// Упакованный канал: подготовка payload -> CommandSeq -> Result -> Ack.
udiGeometryRequest := GVL_HMI.udiGeometryCommandSeq;
xGeometryRequestFresh := FALSE;
IF (udiGeometryRequest <> UDINT#0) AND (udiGeometryRequest <> GVL_HMI.udiGeometryAckSeq) THEN
	stGeometryRequest := GVL_HMI.stGeometryRequest;
	GVL_HMI.uiGeometryResult := UINT#2;
	IF NOT IsHmiCommandFresh(udiIssuedAtMs := GVL_HMI.udiGeometryIssuedAtMs) THEN
		GVL_HMI.uiGeometryResult := UINT#4;
	ELSIF xHmiConnectionAlive THEN
		xGeometryRequestFresh := TRUE;
		IF (stGeometryRequest.uiAction = UINT#8) AND (stGeometryRequest.uiMachine >= UINT#1)
		AND (stGeometryRequest.uiMachine <= UINT#3) THEN
			uiGeometryMachine := stGeometryRequest.uiMachine;
			IF GVL_GEOMETRY_CONTROL.axCallAllowed[uiGeometryMachine] THEN
				IF GVL_GEOMETRY_CONTROL.astCalls[uiGeometryMachine].uiState = UINT#1 THEN
					stGeometryCall := GVL_GEOMETRY_CONTROL.astCalls[uiGeometryMachine];
				ELSE
					GVL_GEOMETRY_CONTROL.udiNextCallId := GVL_GEOMETRY_CONTROL.udiNextCallId + UDINT#1;
					IF GVL_GEOMETRY_CONTROL.udiNextCallId = UDINT#0 THEN GVL_GEOMETRY_CONTROL.udiNextCallId := UDINT#1; END_IF;
					stGeometryCall := stGeometryEmptyCall;
					stGeometryCall.udiId := GVL_GEOMETRY_CONTROL.udiNextCallId;
					stGeometryCall.uiMachine := uiGeometryMachine;
					stGeometryCall.uiProductType := GVL_MULTI_TYPE.Config.auiMachineType[uiGeometryMachine];
				END_IF;
				stGeometryCall.xForced := TRUE; stGeometryCall.uiState := UINT#1;
				GVL_GEOMETRY_CONTROL.astCalls[uiGeometryMachine] := stGeometryCall;
				GVL_GEOMETRY_CONTROL.auiActiveCount[uiGeometryMachine] := UINT#0;
				F_GEOMETRY_EVENT(Call := stGeometryCall); GVL_HMI.uiGeometryResult := UINT#1;
			END_IF;
		ELSIF (stGeometryRequest.uiAction = UINT#12) AND (stGeometryRequest.uiMachine >= UINT#1)
		AND (stGeometryRequest.uiMachine <= UINT#3) THEN
			uiGeometryMachine := stGeometryRequest.uiMachine;
			IF GVL_GEOMETRY_CONTROL.axCancelAllowed[uiGeometryMachine] THEN
				GVL_GEOMETRY_CONTROL.astCalls[uiGeometryMachine].uiState := UINT#6;
				F_GEOMETRY_EVENT(Call := GVL_GEOMETRY_CONTROL.astCalls[uiGeometryMachine]); GVL_HMI.uiGeometryResult := UINT#1;
			END_IF;
		ELSIF (stGeometryRequest.uiAction = UINT#9) AND GVL_GEOMETRY_CONTROL.xAutoChangeAllowed
		AND (stGeometryRequest.udiValue <= UDINT#1) THEN
			GVL_GEOMETRY_CONTROL.xAutoEnabled := stGeometryRequest.udiValue = UDINT#1;
			GVL_HMI.uiGeometryResult := UINT#1;
		ELSIF (stGeometryRequest.uiAction = UINT#10) AND GVL_GEOMETRY_CONTROL.xAutoChangeAllowed
		AND (stGeometryRequest.uiMachine <= UINT#3) AND (stGeometryRequest.udiValue >= UDINT#1)
		AND (stGeometryRequest.udiValue <= UDINT#10000) THEN
			FOR uiGeometryMachine := UINT#1 TO UINT#3 DO
				IF (stGeometryRequest.uiMachine = UINT#0) OR (stGeometryRequest.uiMachine = uiGeometryMachine) THEN
					GVL_GEOMETRY_CONTROL.auiPeriod[uiGeometryMachine] := UDINT_TO_UINT(stGeometryRequest.udiValue);
				END_IF;
			END_FOR;
			GVL_HMI.uiGeometryResult := UINT#1;
		ELSIF (stGeometryRequest.uiAction = UINT#16) AND GVL_GEOMETRY_CONTROL.xSettingsAllowed THEN
			CASE stGeometryRequest.uiMachine OF
				UINT#1: IF stGeometryRequest.udiValue <= UDINT#1 THEN GVL_GEOMETRY_CONTROL.xWaitWhenOccupied := stGeometryRequest.udiValue = UDINT#1; GVL_HMI.uiGeometryResult := UINT#1; END_IF;
				UINT#2: IF (stGeometryRequest.udiValue >= UDINT#100) AND (stGeometryRequest.udiValue <= UDINT#600000) THEN GVL_GEOMETRY_CONTROL.tTransportTimeout := UDINT_TO_TIME(stGeometryRequest.udiValue); GVL_HMI.uiGeometryResult := UINT#1; END_IF;
				UINT#3: IF (stGeometryRequest.udiValue >= UDINT#100) AND (stGeometryRequest.udiValue <= UDINT#60000) THEN GVL_GEOMETRY_CONTROL.tDriveFeedbackTimeout := UDINT_TO_TIME(stGeometryRequest.udiValue); GVL_HMI.uiGeometryResult := UINT#1; END_IF;
				UINT#4: IF (stGeometryRequest.udiValue >= UDINT#100) AND (stGeometryRequest.udiValue <= UDINT#10000) THEN GVL_GEOMETRY_CONTROL.tResetPulse := UDINT_TO_TIME(stGeometryRequest.udiValue); GVL_HMI.uiGeometryResult := UINT#1; END_IF;
				UINT#5: IF (stGeometryRequest.udiValue >= UDINT#1000) AND (stGeometryRequest.udiValue <= UDINT#3600000) THEN GVL_GEOMETRY_CONTROL.tWaitWarningTimeout := UDINT_TO_TIME(stGeometryRequest.udiValue); GVL_HMI.uiGeometryResult := UINT#1; END_IF;
			END_CASE;
		ELSIF (stGeometryRequest.uiStation >= UINT#1) AND (stGeometryRequest.uiStation <= UINT#2) THEN
			uiGeometry := stGeometryRequest.uiStation;
			IF (stGeometryRequest.uiAction >= UINT#1) AND (stGeometryRequest.uiAction <= UINT#7) THEN
				GVL_GEOMETRY_CONTROL.auiAction[uiGeometry] := stGeometryRequest.uiAction;
			ELSIF (stGeometryRequest.uiAction = UINT#11) AND GVL_GEOMETRY_CONTROL.xSupported
			AND GVL_POINT_MANAGER.PointManager.Diag.xXLimitValid
			AND GVL_POINT_MANAGER.PointManager.Diag.xYLimitValid
			AND GVL_POINT_MANAGER.PointManager.Diag.xZLimitValid THEN
				stGeometryConfig := stGeometryRequest.Config;
				stGeometryConfig.lrChangeZ := stGeometryConfig.lrSafeZ;
				xGeometryConfigValid := (stGeometryConfig.lrSpeedFactor >= 0.1) AND (stGeometryConfig.lrSpeedFactor <= 1.0)
					AND (stGeometryConfig.lrSafeZ < 0.0) AND (stGeometryConfig.lrSafeZ >= -10000.0)
					AND (stGeometryConfig.lrX >= GVL_POINT_MANAGER.PointManager.Diag.lrX_MinLimit)
					AND (stGeometryConfig.lrX <= GVL_POINT_MANAGER.PointManager.Diag.lrX_MaxLimit)
					AND (stGeometryConfig.lrY >= GVL_POINT_MANAGER.PointManager.Diag.lrY_MinLimit)
					AND (stGeometryConfig.lrY <= GVL_POINT_MANAGER.PointManager.Diag.lrY_MaxLimit)
					AND (stGeometryConfig.lrZ >= GVL_POINT_MANAGER.PointManager.Diag.lrZ_MinLimit)
					AND (stGeometryConfig.lrZ <= GVL_POINT_MANAGER.PointManager.Diag.lrZ_MaxLimit)
					AND ((stGeometryConfig.lrZ + stGeometryConfig.lrSafeZ) >= GVL_POINT_MANAGER.PointManager.Diag.lrZ_MinLimit);
				IF xGeometryConfigValid THEN
					stGeometryConfig.xConfigured := TRUE;
					IF GVL_CELL_SETTINGS.eTestEnvironment = E_CELL_TEST_ENVIRONMENT.NORMAL THEN GVL_GEOMETRY_CONTROL.astConfig[uiGeometry] := stGeometryConfig;
					ELSE GVL_GEOMETRY_CONTROL.astSimulationConfig[uiGeometry] := stGeometryConfig; END_IF;
					GVL_GEOMETRY_CONTROL.astActiveConfig[uiGeometry] := stGeometryConfig; GVL_HMI.uiGeometryResult := UINT#1;
				END_IF;
			ELSIF (stGeometryRequest.uiAction = UINT#13) AND GVL_GEOMETRY_CONTROL.astStatus[uiGeometry].xPointWriteAllowed
			AND GVL_HMI.xPointEditorCaptureAllowed THEN
				GVL_HMI.stGeometryCapture := GVL_GEOMETRY_CONTROL.astActiveConfig[uiGeometry];
				GVL_HMI.stGeometryCapture.lrX := lrRobotActualX; GVL_HMI.stGeometryCapture.lrY := lrRobotActualY;
				GVL_HMI.stGeometryCapture.lrZ := lrRobotActualZ; GVL_HMI.uiGeometryResult := UINT#1;
			ELSIF ((stGeometryRequest.uiAction = UINT#14) OR (stGeometryRequest.uiAction = UINT#15))
			AND GVL_CELL_SETTINGS.xErrorSimulationEnabled
			AND (GVL_CELL_SETTINGS.eTestEnvironment = E_CELL_TEST_ENVIRONMENT.SIMULATION)
			AND GVL_GEOMETRY_CONTROL.xSupported THEN
				GVL_GEOMETRY_CONTROL.axSimulationAlarm[uiGeometry] := stGeometryRequest.uiAction = UINT#14;
				GVL_HMI.uiGeometryResult := UINT#1;
			END_IF;
		END_IF;
	END_IF;
END_IF;

FOR uiGeometry := UINT#1 TO UINT#2 DO
	xGeometryStopAttempt := FALSE;
	IF (GVL_HMI.audiGeometryStopSeq[uiGeometry] <> UDINT#0)
	AND (GVL_HMI.audiGeometryStopSeq[uiGeometry] <> GVL_HMI.audiGeometryStopAck[uiGeometry]) THEN
		GVL_GEOMETRY_CONTROL.auiAction[uiGeometry] := UINT#6;
		xGeometryStopAttempt := TRUE;
		GVL_HMI.audiGeometryStopAck[uiGeometry] := GVL_HMI.audiGeometryStopSeq[uiGeometry];
	END_IF;
	IF GVL_CELL_SETTINGS.eTestEnvironment <> E_CELL_TEST_ENVIRONMENT.NORMAL THEN
		GEOMETRY_SIM[uiGeometry](xInitialize := xGeometryEnvironmentChanged OR xTestInitializePulse,
			xRun := GEOMETRY[uiGeometry].xRunOutput, xReset := GEOMETRY[uiGeometry].xResetOutput,
			xDeposited := GVL_GEOMETRY_CONTROL.astSignals[uiGeometry].xDeposited,
			udiPartId := GVL_GEOMETRY_CONTROL.astSignals[uiGeometry].Call.udiId,
			xRemove := GEOMETRY[uiGeometry].xSimulationEmptyConfirmed,
			xAlarm := GVL_GEOMETRY_CONTROL.axSimulationAlarm[uiGeometry],
			uiTimeFactor := SEL(GVL_CELL_SETTINGS.xSimulationAccelerationActive, UINT#1, GVL_CELL_SETTINGS.uiSimulationTimeFactorApplied));
		xGeometryDriveAlarm := GEOMETRY_SIM[uiGeometry].xDriveAlarm;
		xGeometryDriveRunning := GEOMETRY_SIM[uiGeometry].xDriveRunning;
		xGeometryPartAtEnd := GEOMETRY_SIM[uiGeometry].xPartAtEnd;
	ELSE
		uiGeometryDi := UINT#81 + (uiGeometry - UINT#1) * UINT#2;
		xGeometryDriveAlarm := xPhysicalNormal AND (GVL_PHYSICAL_IO.xMappingVerified OR axIoForced[uiGeometryDi]) AND axPhysicalRaw[uiGeometryDi];
		xGeometryDriveRunning := xPhysicalNormal AND (GVL_PHYSICAL_IO.xMappingVerified OR axIoForced[uiGeometryDi + UINT#1]) AND axPhysicalRaw[uiGeometryDi + UINT#1];
		xGeometryPartAtEnd := GVL_PHYSICAL_IO.axGkPartAtEnd[uiGeometry];
	END_IF;
	stGeometrySignals := GVL_GEOMETRY_CONTROL.astSignals[uiGeometry];
	// Ручное движение также считается работой с ГК; состояние последней точки
	// удерживает блокировку ленты вплоть до подтверждённого отхода.
	IF uiGeometry = UINT#1 THEN
		stGeometrySignals.xRobotInteraction := stGeometrySignals.xRobotInteraction
			OR (GVL_ROBOT.Status.eCurrentPoint = E_POINT_NAME.GEOMETRY_1_PLACE)
			OR (GVL_ROBOT.Status.eCurrentPoint = E_POINT_NAME.GEOMETRY_1_CHANGE)
			OR (GVL_ROBOT.Status.xBusy AND ((GVL_ROBOT.Command.eSetPoint = E_POINT_NAME.GEOMETRY_1_PLACE)
				OR (GVL_ROBOT.Command.eSetPoint = E_POINT_NAME.GEOMETRY_1_CHANGE)));
	ELSE
		stGeometrySignals.xRobotInteraction := stGeometrySignals.xRobotInteraction
			OR (GVL_ROBOT.Status.eCurrentPoint = E_POINT_NAME.GEOMETRY_2_PLACE)
			OR (GVL_ROBOT.Status.eCurrentPoint = E_POINT_NAME.GEOMETRY_2_CHANGE)
			OR (GVL_ROBOT.Status.xBusy AND ((GVL_ROBOT.Command.eSetPoint = E_POINT_NAME.GEOMETRY_2_PLACE)
				OR (GVL_ROBOT.Command.eSetPoint = E_POINT_NAME.GEOMETRY_2_CHANGE)));
	END_IF;
	GEOMETRY[uiGeometry](xInitialize := xGeometryEnvironmentChanged, uiAction := GVL_GEOMETRY_CONTROL.auiAction[uiGeometry],
		xSupported := GVL_GEOMETRY_CONTROL.xSupported AND ((GVL_CELL_SETTINGS.eTestEnvironment <> E_CELL_TEST_ENVIRONMENT.NORMAL) OR GVL_PHYSICAL_IO.xMappingVerified),
		xSimulation := GVL_CELL_SETTINGS.eTestEnvironment <> E_CELL_TEST_ENVIRONMENT.NORMAL,
		xGlobalError := GVL_CELL_CONTROL.xGlobalError, xManual := GVL_CELL_CONTROL.xManual,
		xCellRunning := GVL_CELL_MANAGER.Status.xRunning, xRobotBusy := GVL_ROBOT.Status.xBusy,
		xMotionBusy := xMotionBusy, xHmiAlive := xHmiConnectionAlive, xIoManual := xIoManualActive,
		xReset := GVL_CELL_CONTROL.xReset, xDriveAlarm := xGeometryDriveAlarm,
		xDriveRunning := xGeometryDriveRunning, xPartAtEnd := xGeometryPartAtEnd,
		rSimulationTravel := GEOMETRY_SIM[uiGeometry].rTravel,
		Signals := stGeometrySignals, Config := GVL_GEOMETRY_CONTROL.astActiveConfig[uiGeometry],
		tTransport := GVL_GEOMETRY_CONTROL.tTransportTimeout, tFeedback := GVL_GEOMETRY_CONTROL.tDriveFeedbackTimeout,
		tResetPulse := GVL_GEOMETRY_CONTROL.tResetPulse,
		uiTimeFactor := SEL(GVL_CELL_SETTINGS.xSimulationAccelerationActive, UINT#1, GVL_CELL_SETTINGS.uiSimulationTimeFactorApplied),
		Memory := GVL_GEOMETRY_CONTROL.astActiveMemory[uiGeometry], Status => GVL_GEOMETRY_CONTROL.astStatus[uiGeometry],
		Warning => GVL_GEOMETRY_CONTROL.astWarning[uiGeometry]);
	GVL_GEOMETRY_CONTROL.astStatus[uiGeometry].xConfigAllowed := GVL_GEOMETRY_CONTROL.astStatus[uiGeometry].xConfigAllowed AND GVL_HMI.xPointEditorSaveAllowed;
	// Только доступность канала данных и лимитов; физическая карта, Home,
	// режим, ошибки, движение и состояние станции не ограничивают SAVE.
	GVL_GEOMETRY_CONTROL.astStatus[uiGeometry].xPointWriteAllowed := GVL_GEOMETRY_CONTROL.xSupported
		AND xHmiConnectionAlive AND GVL_POINT_MANAGER.PointManager.Diag.xXLimitValid
		AND GVL_POINT_MANAGER.PointManager.Diag.xYLimitValid
		AND GVL_POINT_MANAGER.PointManager.Diag.xZLimitValid;
	GVL_GEOMETRY_CONTROL.astStatus[uiGeometry].xSimulationAlarmAllowed := GVL_GEOMETRY_CONTROL.xSupported
		AND (GVL_CELL_SETTINGS.eTestEnvironment = E_CELL_TEST_ENVIRONMENT.SIMULATION)
		AND GVL_CELL_SETTINGS.xErrorSimulationEnabled AND xHmiConnectionAlive;
	IF xGeometryRequestFresh AND NOT xGeometryStopAttempt
	AND (udiGeometryRequest <> UDINT#0) AND (udiGeometryRequest <> GVL_HMI.udiGeometryAckSeq)
	AND (stGeometryRequest.uiStation = uiGeometry) AND (stGeometryRequest.uiAction >= UINT#1) AND (stGeometryRequest.uiAction <= UINT#7) THEN
		IF GEOMETRY[uiGeometry].xCommandAccepted THEN GVL_HMI.uiGeometryResult := UINT#1; END_IF;
	END_IF;
	// Точки ГК независимы от механики/баз палет и от включения магазина.
	IF uiGeometry = UINT#1 THEN eGeometryPlace := E_POINT_NAME.GEOMETRY_1_PLACE; eGeometrySafe := E_POINT_NAME.GEOMETRY_1_SAFE; eGeometryChange := E_POINT_NAME.GEOMETRY_1_CHANGE;
	ELSE eGeometryPlace := E_POINT_NAME.GEOMETRY_2_PLACE; eGeometrySafe := E_POINT_NAME.GEOMETRY_2_SAFE; eGeometryChange := E_POINT_NAME.GEOMETRY_2_CHANGE; END_IF;
	GVL_POINT.Points[eGeometryPlace].X := GVL_GEOMETRY_CONTROL.astActiveConfig[uiGeometry].lrX;
	GVL_POINT.Points[eGeometryPlace].Y := GVL_GEOMETRY_CONTROL.astActiveConfig[uiGeometry].lrY;
	GVL_POINT.Points[eGeometryPlace].Z := GVL_GEOMETRY_CONTROL.astActiveConfig[uiGeometry].lrZ;
	GVL_POINT.Points[eGeometryPlace].MagazineSafeZ := GVL_GEOMETRY_CONTROL.astActiveConfig[uiGeometry].lrSafeZ;
	GVL_POINT.Points[eGeometryPlace].MagazineChangeZ := LREAL#0.0;
	GVL_POINT.Points[eGeometryPlace].SpeedFactor := GVL_GEOMETRY_CONTROL.astActiveConfig[uiGeometry].lrSpeedFactor;
	GVL_POINT.Points[eGeometryPlace].xConfigured := GVL_GEOMETRY_CONTROL.astActiveConfig[uiGeometry].xConfigured;
	GVL_POINT.Points[eGeometrySafe] := GVL_POINT.Points[eGeometryPlace];
	GVL_POINT.Points[eGeometrySafe].Z := GVL_POINT.Points[eGeometryPlace].Z + GVL_GEOMETRY_CONTROL.astActiveConfig[uiGeometry].lrSafeZ;
	GVL_POINT.Points[eGeometryChange] := GVL_POINT.Points[eGeometrySafe]; // Legacy CHANGE совпадает с SAFE_Z
END_FOR;
IF (udiGeometryRequest <> UDINT#0) AND (udiGeometryRequest <> GVL_HMI.udiGeometryAckSeq) THEN
	IF GVL_HMI.uiGeometryResult <> UINT#1 THEN
		GVL_GEOMETRY_CONTROL.stCellWarning.uiCode := UINT#51;
		GVL_GEOMETRY_CONTROL.stCellWarning.udiSequence := GVL_GEOMETRY_CONTROL.stCellWarning.udiSequence + UDINT#1;
	END_IF;
	GVL_HMI.udiGeometryAckSeq := udiGeometryRequest;
END_IF;
END_METHOD

METHOD PRIVATE RunMachines
// Импульсные команды HMI изменяют сохранённое разрешение работы станка.
FOR uiMachine := 1 TO 3 DO
	IF GVL_HMI.axMachineDisable[uiMachine] THEN
		GVL_HMI.axMachineUsed[uiMachine] := FALSE;
	ELSIF GVL_HMI.axMachineEnable[uiMachine] AND axMachinePointsReady[uiMachine] THEN
		GVL_HMI.axMachineUsed[uiMachine] := TRUE;
	END_IF;
END_FOR;


MACHINE_1.stPoints.eAbove := E_POINT_NAME.MACHINE_1_ABOVE;
MACHINE_1.stPoints.eChuck := E_POINT_NAME.MACHINE_1_CHUCK_POSITION;
MACHINE_1.stPoints.eChuckApproach := E_POINT_NAME.MACHINE_1_CHUCK_APROACH;
MACHINE_1.stPoints.eInside := E_POINT_NAME.MACHINE_1_INSIDE;
MACHINE_1.stPoints.eNone := E_POINT_NAME.NONE;

// NORMAL получает только физическую обратную связь; обе тестовые среды — модель.
IF GVL_CELL_SETTINGS.eTestEnvironment <> E_CELL_TEST_ENVIRONMENT.NORMAL THEN
// Виртуальные устройства исполняют команду предыдущего цикла. Затем слой
// инъекции формирует обратную связь, которую увидит технологический автомат.
MACHINE_1_SIM(
	xTestInitialize := xTestInitializePulse OR xTestAbortActive,
	uiTestInitialState := GVL_HMI.stTestScenario.auiMachineState[1],
	xSafetyDoorOpen := GVL_CELL_SETTINGS.xErrorSimulationEnabled
		AND GVL_HMI.axMachineSimSafetyDoorOpen[1],
	Command := GVL_MACHINE.Command[1].stIo,
	FaultRequest := astMachineFaultRequest[1],
	xSimulationAccelerationEnable := GVL_CELL_SETTINGS.xSimulationAccelerationActive,
	uiSimulationTimeFactor := GVL_CELL_SETTINGS.uiSimulationTimeFactorApplied,
	tDoorOpenTime := GVL_HMI.tMachineDoorOpenTime,
	tDoorCloseTime := GVL_HMI.tMachineDoorCloseTime,
	tChuckOpenTime := GVL_HMI.tMachineChuckOpenTime,
	tChuckCloseTime := GVL_HMI.tMachineChuckCloseTime,
	tCycleTime := GVL_HMI.tMachineCycleTime[1]
);
MACHINE_2_SIM(
	xTestInitialize := xTestInitializePulse OR xTestAbortActive,
	uiTestInitialState := GVL_HMI.stTestScenario.auiMachineState[2],
	xSafetyDoorOpen := GVL_CELL_SETTINGS.xErrorSimulationEnabled
		AND GVL_HMI.axMachineSimSafetyDoorOpen[2],
	Command := GVL_MACHINE.Command[2].stIo,
	FaultRequest := astMachineFaultRequest[2],
	xSimulationAccelerationEnable := GVL_CELL_SETTINGS.xSimulationAccelerationActive,
	uiSimulationTimeFactor := GVL_CELL_SETTINGS.uiSimulationTimeFactorApplied,
	tDoorOpenTime := GVL_HMI.tMachineDoorOpenTime,
	tDoorCloseTime := GVL_HMI.tMachineDoorCloseTime,
	tChuckOpenTime := GVL_HMI.tMachineChuckOpenTime,
	tChuckCloseTime := GVL_HMI.tMachineChuckCloseTime,
	tCycleTime := GVL_HMI.tMachineCycleTime[2]
);
MACHINE_3_SIM(
	xTestInitialize := xTestInitializePulse OR xTestAbortActive,
	uiTestInitialState := GVL_HMI.stTestScenario.auiMachineState[3],
	xSafetyDoorOpen := GVL_CELL_SETTINGS.xErrorSimulationEnabled
		AND GVL_HMI.axMachineSimSafetyDoorOpen[3],
	Command := GVL_MACHINE.Command[3].stIo,
	FaultRequest := astMachineFaultRequest[3],
	xSimulationAccelerationEnable := GVL_CELL_SETTINGS.xSimulationAccelerationActive,
	uiSimulationTimeFactor := GVL_CELL_SETTINGS.uiSimulationTimeFactorApplied,
	tDoorOpenTime := GVL_HMI.tMachineDoorOpenTime,
	tDoorCloseTime := GVL_HMI.tMachineDoorCloseTime,
	tChuckOpenTime := GVL_HMI.tMachineChuckOpenTime,
	tChuckCloseTime := GVL_HMI.tMachineChuckCloseTime,
	tCycleTime := GVL_HMI.tMachineCycleTime[3]
);

END_IF;
IF GVL_CELL_SETTINGS.eTestEnvironment = E_CELL_TEST_ENVIRONMENT.NORMAL THEN
	astMachineStatusRaw := GVL_MACHINE.astPhysicalInput;
ELSE
	astMachineStatusRaw[1] := MACHINE_1_SIM.Status;
	astMachineStatusRaw[2] := MACHINE_2_SIM.Status;
	astMachineStatusRaw[3] := MACHINE_3_SIM.Status;
END_IF;

MACHINE_1_FAULT(
	Request := astMachineFaultRequest[1],
	MachineStatusRaw := astMachineStatusRaw[1],
	RobotStatusRaw := GVL_ROBOT.Status,
	NominalTimeouts := GVL_CELL_SETTINGS.stMachineTimeouts
);
MACHINE_2_FAULT(
	Request := astMachineFaultRequest[2],
	MachineStatusRaw := astMachineStatusRaw[2],
	RobotStatusRaw := GVL_ROBOT.Status,
	NominalTimeouts := GVL_CELL_SETTINGS.stMachineTimeouts
);
MACHINE_3_FAULT(
	Request := astMachineFaultRequest[3],
	MachineStatusRaw := astMachineStatusRaw[3],
	RobotStatusRaw := GVL_ROBOT.Status,
	NominalTimeouts := GVL_CELL_SETTINGS.stMachineTimeouts
);

MACHINE_1(
	xTestInitialize := xTestInitializePulse OR xTestAbortActive,
	uiTestInitialState := GVL_HMI.stTestScenario.auiMachineState[1],
	uiTestProductType := GVL_HMI.stTestScenario.auiMachineType[1],
	xExecute := GVL_CELL_MANAGER.Command.axMachineExecute[1],
	xReset := GVL_HMI.axMachineReset[1],
	xResetGlobal := GVL_CELL_CONTROL.xReset,
	xGlobalError := GVL_CELL_CONTROL.xGlobalError,
	xManualMode := GVL_CELL_CONTROL.xManual,
	xIoManual := xIoManualActive,
	xAutomaticUseEnabled := GVL_HMI.axMachineUsed[1],
	xPointsConfigured := axMachinePointsReady[1],
	xSafetyDoorControlEnabled := GVL_CELL_SETTINGS.eTestEnvironment <> E_CELL_TEST_ENVIRONMENT.NORMAL,
	xHmiOpenSafetyDoor := GVL_HMI.axMachineManualSafetyDoorOpen[1],
	xHmiCloseSafetyDoor := GVL_HMI.axMachineManualSafetyDoorClose[1],
	xHmiOpenHatch := GVL_HMI.axMachineManualHatchOpen[1],
	xHmiCloseHatch := GVL_HMI.axMachineManualHatchClose[1],
	xHmiUnlockHatch := GVL_HMI.axMachineManualHatchUnlock[1],
	xHmiLockHatch := GVL_HMI.axMachineManualHatchLock[1],
	xHmiOpenChuck := GVL_HMI.axMachineManualChuckOpen[1],
	xHmiCloseChuck := GVL_HMI.axMachineManualChuckClose[1],
	xHmiEnable := GVL_HMI.axMachineEnable[1],
	xHmiDisable := GVL_HMI.axMachineDisable[1],
	xHmiSetBlank := GVL_HMI.axMachineSetBlank[1],
	xHmiSetDetail := GVL_HMI.axMachineSetDetail[1],
	xHmiAcceptDoor := GVL_HMI.axMachineAcceptDoor[1],
	xHmiRejectDoor := GVL_HMI.axMachineRejectDoor[1],
	xHmiAcceptRunCNC := GVL_HMI.axMachineAcceptRun[1],
	xHmiRejectRunCNC := GVL_HMI.axMachineRejectRun[1],
	xUseHmiCycleTime := GVL_HMI.xUseHmiCycleTime[1],
	tHmiCycleTime := GVL_HMI.tMachineCycleTime[1],
	stTimeouts := MACHINE_1_FAULT.Timeouts,
	stChangeRecipe := GVL_CELL_SETTINGS.CHANGE_MACHINE,
	stLoadRecipe := GVL_CELL_SETTINGS.LOAD_MACHINE,
	stUnloadRecipe := GVL_CELL_SETTINGS.UNLOAD_MACHINE,
	stMachineStatus := MACHINE_1_FAULT.MachineStatus,
	stRobotStatus := MACHINE_1_FAULT.RobotStatus,
	eRobotTargetPoint := GVL_ROBOT.Diag.eActivePoint,
	xRobotMotionBusy := xMotionBusy,
	Command => GVL_MACHINE.Command[1],
	Status => GVL_MACHINE.Status[1],
	Diag => GVL_MACHINE.Diag[1],
	Error => GVL_MACHINE.Error[1]
);

MACHINE_2.stPoints.eAbove := E_POINT_NAME.MACHINE_2_ABOVE;
MACHINE_2.stPoints.eChuck := E_POINT_NAME.MACHINE_2_CHUCK_POSITION;
MACHINE_2.stPoints.eChuckApproach := E_POINT_NAME.MACHINE_2_CHUCK_APROACH;
MACHINE_2.stPoints.eInside := E_POINT_NAME.MACHINE_2_INSIDE;
MACHINE_2.stPoints.eNone := E_POINT_NAME.NONE;

MACHINE_2(
	xTestInitialize := xTestInitializePulse OR xTestAbortActive,
	uiTestInitialState := GVL_HMI.stTestScenario.auiMachineState[2],
	uiTestProductType := GVL_HMI.stTestScenario.auiMachineType[2],
	xExecute := GVL_CELL_MANAGER.Command.axMachineExecute[2],
	xReset := GVL_HMI.axMachineReset[2],
	xResetGlobal := GVL_CELL_CONTROL.xReset,
	xGlobalError := GVL_CELL_CONTROL.xGlobalError,
	xManualMode := GVL_CELL_CONTROL.xManual,
	xIoManual := xIoManualActive,
	xAutomaticUseEnabled := GVL_HMI.axMachineUsed[2],
	xPointsConfigured := axMachinePointsReady[2],
	xSafetyDoorControlEnabled := GVL_CELL_SETTINGS.eTestEnvironment <> E_CELL_TEST_ENVIRONMENT.NORMAL,
	xHmiOpenSafetyDoor := GVL_HMI.axMachineManualSafetyDoorOpen[2],
	xHmiCloseSafetyDoor := GVL_HMI.axMachineManualSafetyDoorClose[2],
	xHmiOpenHatch := GVL_HMI.axMachineManualHatchOpen[2],
	xHmiCloseHatch := GVL_HMI.axMachineManualHatchClose[2],
	xHmiUnlockHatch := GVL_HMI.axMachineManualHatchUnlock[2],
	xHmiLockHatch := GVL_HMI.axMachineManualHatchLock[2],
	xHmiOpenChuck := GVL_HMI.axMachineManualChuckOpen[2],
	xHmiCloseChuck := GVL_HMI.axMachineManualChuckClose[2],
	xHmiEnable := GVL_HMI.axMachineEnable[2],
	xHmiDisable := GVL_HMI.axMachineDisable[2],
	xHmiSetBlank := GVL_HMI.axMachineSetBlank[2],
	xHmiSetDetail := GVL_HMI.axMachineSetDetail[2],
	xHmiAcceptDoor := GVL_HMI.axMachineAcceptDoor[2],
	xHmiRejectDoor := GVL_HMI.axMachineRejectDoor[2],
	xHmiAcceptRunCNC := GVL_HMI.axMachineAcceptRun[2],
	xHmiRejectRunCNC := GVL_HMI.axMachineRejectRun[2],
	xUseHmiCycleTime := GVL_HMI.xUseHmiCycleTime[2],
	tHmiCycleTime := GVL_HMI.tMachineCycleTime[2],
	stTimeouts := MACHINE_2_FAULT.Timeouts,
	stChangeRecipe := GVL_CELL_SETTINGS.CHANGE_MACHINE,
	stLoadRecipe := GVL_CELL_SETTINGS.LOAD_MACHINE,
	stUnloadRecipe := GVL_CELL_SETTINGS.UNLOAD_MACHINE,
	stMachineStatus := MACHINE_2_FAULT.MachineStatus,
	stRobotStatus := MACHINE_2_FAULT.RobotStatus,
	eRobotTargetPoint := GVL_ROBOT.Diag.eActivePoint,
	xRobotMotionBusy := xMotionBusy,
	Command => GVL_MACHINE.Command[2],
	Status => GVL_MACHINE.Status[2],
	Diag => GVL_MACHINE.Diag[2],
	Error => GVL_MACHINE.Error[2]
);

MACHINE_3.stPoints.eAbove := E_POINT_NAME.MACHINE_3_ABOVE;
MACHINE_3.stPoints.eChuck := E_POINT_NAME.MACHINE_3_CHUCK_POSITION;
MACHINE_3.stPoints.eChuckApproach := E_POINT_NAME.MACHINE_3_CHUCK_APROACH;
MACHINE_3.stPoints.eInside := E_POINT_NAME.MACHINE_3_INSIDE;
MACHINE_3.stPoints.eNone := E_POINT_NAME.NONE;

MACHINE_3(
	xTestInitialize := xTestInitializePulse OR xTestAbortActive,
	uiTestInitialState := GVL_HMI.stTestScenario.auiMachineState[3],
	uiTestProductType := GVL_HMI.stTestScenario.auiMachineType[3],
	xExecute := GVL_CELL_MANAGER.Command.axMachineExecute[3],
	xReset := GVL_HMI.axMachineReset[3],
	xResetGlobal := GVL_CELL_CONTROL.xReset,
	xGlobalError := GVL_CELL_CONTROL.xGlobalError,
	xManualMode := GVL_CELL_CONTROL.xManual,
	xIoManual := xIoManualActive,
	xAutomaticUseEnabled := GVL_HMI.axMachineUsed[3],
	xPointsConfigured := axMachinePointsReady[3],
	xSafetyDoorControlEnabled := GVL_CELL_SETTINGS.eTestEnvironment <> E_CELL_TEST_ENVIRONMENT.NORMAL,
	xHmiOpenSafetyDoor := GVL_HMI.axMachineManualSafetyDoorOpen[3],
	xHmiCloseSafetyDoor := GVL_HMI.axMachineManualSafetyDoorClose[3],
	xHmiOpenHatch := GVL_HMI.axMachineManualHatchOpen[3],
	xHmiCloseHatch := GVL_HMI.axMachineManualHatchClose[3],
	xHmiUnlockHatch := GVL_HMI.axMachineManualHatchUnlock[3],
	xHmiLockHatch := GVL_HMI.axMachineManualHatchLock[3],
	xHmiOpenChuck := GVL_HMI.axMachineManualChuckOpen[3],
	xHmiCloseChuck := GVL_HMI.axMachineManualChuckClose[3],
	xHmiEnable := GVL_HMI.axMachineEnable[3],
	xHmiDisable := GVL_HMI.axMachineDisable[3],
	xHmiSetBlank := GVL_HMI.axMachineSetBlank[3],
	xHmiSetDetail := GVL_HMI.axMachineSetDetail[3],
	xHmiAcceptDoor := GVL_HMI.axMachineAcceptDoor[3],
	xHmiRejectDoor := GVL_HMI.axMachineRejectDoor[3],
	xHmiAcceptRunCNC := GVL_HMI.axMachineAcceptRun[3],
	xHmiRejectRunCNC := GVL_HMI.axMachineRejectRun[3],
	xUseHmiCycleTime := GVL_HMI.xUseHmiCycleTime[3],
	tHmiCycleTime := GVL_HMI.tMachineCycleTime[3],
	stTimeouts := MACHINE_3_FAULT.Timeouts,
	stChangeRecipe := GVL_CELL_SETTINGS.CHANGE_MACHINE,
	stLoadRecipe := GVL_CELL_SETTINGS.LOAD_MACHINE,
	stUnloadRecipe := GVL_CELL_SETTINGS.UNLOAD_MACHINE,
	stMachineStatus := MACHINE_3_FAULT.MachineStatus,
	stRobotStatus := MACHINE_3_FAULT.RobotStatus,
	eRobotTargetPoint := GVL_ROBOT.Diag.eActivePoint,
	xRobotMotionBusy := xMotionBusy,
	Command => GVL_MACHINE.Command[3],
	Status => GVL_MACHINE.Status[3],
	Diag => GVL_MACHINE.Diag[3],
	Error => GVL_MACHINE.Error[3]
);

// Публичный IO-снимок совпадает с обратной связью, которую анализирует FB_MACHINE.
GVL_MACHINE.Status[1].stIo := MACHINE_1_FAULT.MachineStatus;
GVL_MACHINE.Status[2].stIo := MACHINE_2_FAULT.MachineStatus;
GVL_MACHINE.Status[3].stIo := MACHINE_3_FAULT.MachineStatus;
END_METHOD

METHOD PRIVATE ApplyIoOutputOverrides
// Прямой ручной режим владеет всеми DO. Штатные уровни остаются отдельно для возврата программе.
axIoAutoDo[1] := GVL_PHYSICAL_IO.xDoMachine1HatchClosed;
axIoAutoDo[2] := GVL_PHYSICAL_IO.xDoMachine1HatchUnLock;
axIoAutoDo[3] := GVL_PHYSICAL_IO.xDoMachine1ClampChuck;
axIoAutoDo[4] := GVL_PHYSICAL_IO.xDoMachine1UnclampChuck;
axIoAutoDo[5] := GVL_PHYSICAL_IO.xDoMachine1StartCycle;
axIoAutoDo[6] := GVL_PHYSICAL_IO.xDoMachine2HatchClosed;
axIoAutoDo[7] := GVL_PHYSICAL_IO.xDoMachine2HatchUnLock;
axIoAutoDo[8] := GVL_PHYSICAL_IO.xDoMachine2ClampChuck;
axIoAutoDo[9] := GVL_PHYSICAL_IO.xDoMachine2UnclampChuck;
axIoAutoDo[10] := GVL_PHYSICAL_IO.xDoMachine2StartCycle;
axIoAutoDo[11] := GVL_PHYSICAL_IO.xDoMachine3HatchClosed;
axIoAutoDo[12] := GVL_PHYSICAL_IO.xDoMachine3HatchUnLock;
axIoAutoDo[13] := GVL_PHYSICAL_IO.xDoMachine3ClampChuck;
axIoAutoDo[14] := GVL_PHYSICAL_IO.xDoMachine3UnclampChuck;
axIoAutoDo[15] := GVL_PHYSICAL_IO.xDoMachine3StartCycle;
axIoAutoDo[16] := GVL_PHYSICAL_IO.xDoGripper1Open;
axIoAutoDo[17] := GVL_PHYSICAL_IO.xDoGripper2Open;
axIoAutoDo[18] := GVL_PHYSICAL_IO.xDoRotateToDetail;
axIoAutoDo[19] := GVL_PHYSICAL_IO.xDoDoor1Unlock;
axIoAutoDo[20] := GVL_PHYSICAL_IO.xDoDoor2Unlock;
axIoAutoDo[21] := GVL_PHYSICAL_IO.xDoDoor3Unlock;
axIoAutoDo[22] := GVL_PHYSICAL_IO.xDoDoor4Unlock;
axIoAutoDo[23] := GVL_PHYSICAL_IO.xDoSafetyRelayReset;
axIoAutoDo[24] := GVL_PHYSICAL_IO.xDoSignalTowerGreenOutput;
axIoAutoDo[25] := GVL_PHYSICAL_IO.xDoSignalTowerAmberOutput;
axIoAutoDo[26] := GVL_PHYSICAL_IO.xDoSignalTowerRedOutput;
axIoAutoDo[27] := GVL_PHYSICAL_IO.xDoDoor1ButtonLamp;
axIoAutoDo[28] := GVL_PHYSICAL_IO.xDoDoor2ButtonLamp;
axIoAutoDo[29] := GVL_PHYSICAL_IO.xDoDoor3ButtonLamp;
axIoAutoDo[30] := GVL_PHYSICAL_IO.xDoDoor4ButtonLamp;
axIoAutoDo[31] := GVL_PHYSICAL_IO.xDoMagazine1LockIn;
axIoAutoDo[32] := GVL_PHYSICAL_IO.xDoMagazine1LockOut;
axIoAutoDo[33] := GVL_PHYSICAL_IO.xDoMagazine1StopIn;
axIoAutoDo[34] := GVL_PHYSICAL_IO.xDoMagazine1StopOut;
axIoAutoDo[35] := GVL_PHYSICAL_IO.xDoMagazine1LiftUp;
axIoAutoDo[36] := GVL_PHYSICAL_IO.xDoMagazine1LiftDown;
axIoAutoDo[37] := FALSE; // Удалённый сигнал; индекс журнала не переиспользовать.
axIoAutoDo[38] := FALSE; // Удалённый сигнал; индекс журнала не переиспользовать.
axIoAutoDo[39] := FALSE; // Удалённый сигнал; индекс журнала не переиспользовать.
axIoAutoDo[40] := GVL_PHYSICAL_IO.xDoCellAlarmHorn;
axIoAutoDo[41] := GVL_PHYSICAL_IO.xDoGk1DriveRun;
axIoAutoDo[42] := GVL_PHYSICAL_IO.xDoGk1DriveReset;
axIoAutoDo[43] := GVL_PHYSICAL_IO.xDoMagazine2LockIn;
axIoAutoDo[44] := GVL_PHYSICAL_IO.xDoMagazine2LockOut;
axIoAutoDo[45] := GVL_PHYSICAL_IO.xDoMagazine2StopIn;
axIoAutoDo[46] := GVL_PHYSICAL_IO.xDoMagazine2StopOut;
axIoAutoDo[47] := GVL_PHYSICAL_IO.xDoMagazine2LiftUp;
axIoAutoDo[48] := GVL_PHYSICAL_IO.xDoMagazine2LiftDown;
axIoAutoDo[49] := GVL_PHYSICAL_IO.xDoGk2DriveRun;
axIoAutoDo[50] := GVL_PHYSICAL_IO.xDoGk2DriveReset;
IF xIoManualActive AND NOT GVL_CELL_CONTROL.xManual THEN xIoManualActive := FALSE; END_IF;
GVL_HMI.xIoManualControlActive := xIoManualActive;
GVL_HMI.xIoDoOverrideAllowed := xIoManualActive AND GVL_CELL_CONTROL.xManual;
GVL_HMI.uiIoDoBlockReason := GVL_HMI.uiIoOverrideBlockReason;
IF GVL_HMI.xIoDoOverrideAllowed THEN GVL_HMI.uiIoDoBlockReason := UINT#0; END_IF;

FOR uiIoIndex := UINT#1 TO UINT#50 DO
    // 37..39 удалены из каталога; остальные индексы сохраняют смысл старых событий.
    IF (uiIoIndex >= UINT#37) AND (uiIoIndex <= UINT#39) THEN
        axIoDoForced[uiIoIndex] := FALSE;
        axIoDoForceValue[uiIoIndex] := FALSE;
    END_IF;
    axIoDoAllowed[uiIoIndex] := GVL_HMI.xIoDoOverrideAllowed AND ((uiIoIndex < UINT#37) OR (uiIoIndex > UINT#39));
    axIoDoOnAllowed[uiIoIndex] := axIoDoAllowed[uiIoIndex]; // Совместимость транспорта: включение и отключение равноправны.
    axIoDoInhibited[uiIoIndex] := FALSE; // Старый механизм блокировки снят.
    IF NOT xIoManualActive AND axIoDoForced[uiIoIndex] THEN
        IF xIoManualEndedByOperator THEN
            AppendIoEvent(usiDirection := USINT#2, uiIndex := uiIoIndex, usiKind := USINT#8,
                xOld := axIoDoForceValue[uiIoIndex], xNew := axIoAutoDo[uiIoIndex]);
        ELSE
            AppendIoEvent(usiDirection := USINT#2, uiIndex := uiIoIndex, usiKind := USINT#9,
                xOld := axIoDoForceValue[uiIoIndex], xNew := axIoAutoDo[uiIoIndex]);
        END_IF;
        axIoDoForced[uiIoIndex] := FALSE;
    END_IF;
END_FOR;

xIoDoRejected := FALSE;
udiIoRequestSeq := GVL_HMI.udiIoOverrideCommandSeq;
uiIoRequestAction := GVL_HMI.uiIoOverrideAction;
uiIoRequestIndex := GVL_HMI.uiIoOverrideIndex;
xIoRequestValue := GVL_HMI.xIoOverrideValue;
IF (udiIoRequestSeq <> GVL_HMI.udiIoOverrideAckSeq) AND (uiIoRequestAction >= UINT#4) AND (uiIoRequestAction <= UINT#9) THEN
    IF uiIoRequestAction <= UINT#6 THEN
        GVL_HMI.uiIoOverrideResult := UINT#3;
        IF NOT IsHmiCommandFresh(udiIssuedAtMs := GVL_HMI.udiIoOverrideIssuedAtMs) THEN
            GVL_HMI.uiIoOverrideResult := UINT#4;
        ELSIF uiIoRequestAction = UINT#6 THEN
            FOR uiIoIndex := UINT#1 TO UINT#50 DO
                IF axIoDoForced[uiIoIndex] THEN
                    AppendIoEvent(usiDirection := USINT#2, uiIndex := uiIoIndex, usiKind := USINT#8,
                        xOld := axIoDoForceValue[uiIoIndex], xNew := axIoAutoDo[uiIoIndex]);
                END_IF;
                axIoDoForceValue[uiIoIndex] := axIoAutoDo[uiIoIndex];
                axIoDoForced[uiIoIndex] := FALSE;
            END_FOR;
            GVL_HMI.uiIoOverrideResult := UINT#1;
        ELSIF (uiIoRequestIndex >= UINT#1) AND (uiIoRequestIndex <= UINT#50) AND ((uiIoRequestIndex < UINT#37) OR (uiIoRequestIndex > UINT#39)) THEN
            IF uiIoRequestAction = UINT#5 THEN
                IF axIoDoForced[uiIoRequestIndex] THEN
                    AppendIoEvent(usiDirection := USINT#2, uiIndex := uiIoRequestIndex, usiKind := USINT#8,
                        xOld := axIoDoForceValue[uiIoRequestIndex], xNew := axIoAutoDo[uiIoRequestIndex]);
                END_IF;
                axIoDoForceValue[uiIoRequestIndex] := axIoAutoDo[uiIoRequestIndex];
                axIoDoForced[uiIoRequestIndex] := FALSE;
                GVL_HMI.uiIoOverrideResult := UINT#1;
            ELSIF GVL_HMI.xIoDoOverrideAllowed THEN
                IF NOT axIoDoForced[uiIoRequestIndex] OR (axIoDoForceValue[uiIoRequestIndex] <> xIoRequestValue) THEN
                    AppendIoEvent(usiDirection := USINT#2, uiIndex := uiIoRequestIndex, usiKind := USINT#7,
                        xOld := axIoOutput[uiIoRequestIndex], xNew := xIoRequestValue);
                END_IF;
                axIoDoForced[uiIoRequestIndex] := TRUE;
                axIoDoForceValue[uiIoRequestIndex] := xIoRequestValue;
                IF (uiIoRequestIndex >= UINT#31) AND (uiIoRequestIndex <= UINT#36) THEN axIoMagazineInvalidated[1] := TRUE;
                ELSIF (uiIoRequestIndex >= UINT#43) AND (uiIoRequestIndex <= UINT#48) THEN axIoMagazineInvalidated[2] := TRUE;
                END_IF;
                GVL_HMI.uiIoOverrideResult := UINT#1;
            ELSE
                GVL_HMI.uiIoOverrideResult := UINT#2;
            END_IF;
        END_IF;
    END_IF;
    xIoDoRejected := GVL_HMI.uiIoOverrideResult <> UINT#1;
    GVL_HMI.udiIoOverrideAckSeq := udiIoRequestSeq;
END_IF;

// Намеренно без Safety, пар катушек, режима Modbus, импульсных ограничений и технологических FB.
IF xIoManualActive THEN
    GVL_PHYSICAL_IO.xDoMachine1HatchClosed := axIoDoForceValue[1];
    GVL_PHYSICAL_IO.xDoMachine1HatchUnLock := axIoDoForceValue[2];
    GVL_PHYSICAL_IO.xDoMachine1ClampChuck := axIoDoForceValue[3];
    GVL_PHYSICAL_IO.xDoMachine1UnclampChuck := axIoDoForceValue[4];
    GVL_PHYSICAL_IO.xDoMachine1StartCycle := axIoDoForceValue[5];
    GVL_PHYSICAL_IO.xDoMachine2HatchClosed := axIoDoForceValue[6];
    GVL_PHYSICAL_IO.xDoMachine2HatchUnLock := axIoDoForceValue[7];
    GVL_PHYSICAL_IO.xDoMachine2ClampChuck := axIoDoForceValue[8];
    GVL_PHYSICAL_IO.xDoMachine2UnclampChuck := axIoDoForceValue[9];
    GVL_PHYSICAL_IO.xDoMachine2StartCycle := axIoDoForceValue[10];
    GVL_PHYSICAL_IO.xDoMachine3HatchClosed := axIoDoForceValue[11];
    GVL_PHYSICAL_IO.xDoMachine3HatchUnLock := axIoDoForceValue[12];
    GVL_PHYSICAL_IO.xDoMachine3ClampChuck := axIoDoForceValue[13];
    GVL_PHYSICAL_IO.xDoMachine3UnclampChuck := axIoDoForceValue[14];
    GVL_PHYSICAL_IO.xDoMachine3StartCycle := axIoDoForceValue[15];
    GVL_PHYSICAL_IO.xDoGripper1Open := axIoDoForceValue[16];
    GVL_PHYSICAL_IO.xDoGripper2Open := axIoDoForceValue[17];
    GVL_PHYSICAL_IO.xDoRotateToDetail := axIoDoForceValue[18];
    GVL_PHYSICAL_IO.xDoDoor1Unlock := axIoDoForceValue[19];
    GVL_PHYSICAL_IO.xDoDoor2Unlock := axIoDoForceValue[20];
    GVL_PHYSICAL_IO.xDoDoor3Unlock := axIoDoForceValue[21];
    GVL_PHYSICAL_IO.xDoDoor4Unlock := axIoDoForceValue[22];
    GVL_PHYSICAL_IO.xDoSafetyRelayReset := axIoDoForceValue[23];
    GVL_PHYSICAL_IO.xDoSignalTowerGreenOutput := axIoDoForceValue[24];
    GVL_PHYSICAL_IO.xDoSignalTowerAmberOutput := axIoDoForceValue[25];
    GVL_PHYSICAL_IO.xDoSignalTowerRedOutput := axIoDoForceValue[26];
    GVL_PHYSICAL_IO.xDoDoor1ButtonLamp := axIoDoForceValue[27];
    GVL_PHYSICAL_IO.xDoDoor2ButtonLamp := axIoDoForceValue[28];
    GVL_PHYSICAL_IO.xDoDoor3ButtonLamp := axIoDoForceValue[29];
    GVL_PHYSICAL_IO.xDoDoor4ButtonLamp := axIoDoForceValue[30];
    GVL_PHYSICAL_IO.xDoMagazine1LockIn := axIoDoForceValue[31];
    GVL_PHYSICAL_IO.xDoMagazine1LockOut := axIoDoForceValue[32];
    GVL_PHYSICAL_IO.xDoMagazine1StopIn := axIoDoForceValue[33];
    GVL_PHYSICAL_IO.xDoMagazine1StopOut := axIoDoForceValue[34];
    GVL_PHYSICAL_IO.xDoMagazine1LiftUp := axIoDoForceValue[35];
    GVL_PHYSICAL_IO.xDoMagazine1LiftDown := axIoDoForceValue[36];
    GVL_PHYSICAL_IO.xDoCellAlarmHorn := axIoDoForceValue[40];
    GVL_PHYSICAL_IO.xDoGk1DriveRun := axIoDoForceValue[41];
    GVL_PHYSICAL_IO.xDoGk1DriveReset := axIoDoForceValue[42];
    GVL_PHYSICAL_IO.xDoMagazine2LockIn := axIoDoForceValue[43];
    GVL_PHYSICAL_IO.xDoMagazine2LockOut := axIoDoForceValue[44];
    GVL_PHYSICAL_IO.xDoMagazine2StopIn := axIoDoForceValue[45];
    GVL_PHYSICAL_IO.xDoMagazine2StopOut := axIoDoForceValue[46];
    GVL_PHYSICAL_IO.xDoMagazine2LiftUp := axIoDoForceValue[47];
    GVL_PHYSICAL_IO.xDoMagazine2LiftDown := axIoDoForceValue[48];
    GVL_PHYSICAL_IO.xDoGk2DriveRun := axIoDoForceValue[49];
    GVL_PHYSICAL_IO.xDoGk2DriveReset := axIoDoForceValue[50];
END_IF;
END_METHOD

METHOD PRIVATE RunAlarms
// Единая кнопка подсвечивается только тогда, когда существует хотя бы одна авария
// и каждый активный владелец общей команды готов принять тот же импульс сброса.
// Диагностические защёлки симуляторов станков сюда не входят: они обслуживаются
// отдельной командой «Сброс симулятора» на экране инъекций.
xAlarmResetRequired := (GVL_GEOMETRY_CONTROL.xSupported AND (GVL_GEOMETRY_CONTROL.astStatus[1].xError
	OR GVL_GEOMETRY_CONTROL.astStatus[2].xError))
	OR GVL_CELL_MANAGER.Status.xError
	OR (CELL_SAFETY.Error.dwAlarmActive <> DWORD#0)
	OR GVL_ROBOT.Status.xError
	OR GVL_MACHINE.Status[1].xError
	OR GVL_MACHINE.Status[2].xError
	OR GVL_MACHINE.Status[3].xError
	OR GVL_MAGAZINE.astStatus[1].xError
	OR GVL_MAGAZINE.astStatus[2].xError
	OR (NOT GVL_HMI.xModbusMode AND GVL_AXIS.arrAxis[1].Status.xError)
	OR (NOT GVL_HMI.xModbusMode AND GVL_AXIS.arrAxis[2].Status.xError)
	OR (NOT GVL_HMI.xModbusMode AND GVL_AXIS.arrAxis[3].Status.xError)
	OR (NOT GVL_HMI.xModbusMode AND GVL_AXIS_GROUP.AxisGroup.Status.xLocalError)
	OR (NOT GVL_HMI.xModbusMode AND GVL_AXIS_GROUP.AxisGroup.Status.xLogicalError)
	OR (NOT GVL_HMI.xModbusMode AND GVL_AXIS_GROUP.AxisGroup.Status.xGroupError)
	OR (NOT GVL_HMI.xModbusMode AND (GVL_MOTION_MANAGER.stMotionManager.Error.dwAlarmActive <> DWORD#0))
	OR (NOT GVL_HMI.xModbusMode AND (GVL_POINT_MANAGER.PointManager.Error.dwAlarmActive <> DWORD#0))
	OR (NOT GVL_HMI.xModbusMode AND (GVL_ROBOT.GripperError.dwAlarmActive <> DWORD#0));

xAlarmResetAllowed := ((GVL_TWO_PALLET.uiMode = 0) OR ((NOT GVL_TWO_PALLET.astStatus[1].xError OR GVL_TWO_PALLET.astStatus[1].xResetAllowed) AND (NOT GVL_TWO_PALLET.astStatus[2].xError OR GVL_TWO_PALLET.astStatus[2].xResetAllowed))) AND xAlarmResetRequired
	AND (CELL_SAFETY.Error.dwAlarmActive = DWORD#0)
	AND (NOT GVL_GEOMETRY_CONTROL.xSupported OR NOT GVL_GEOMETRY_CONTROL.astStatus[1].xError OR GVL_GEOMETRY_CONTROL.astStatus[1].xResetAllowed)
	AND (NOT GVL_GEOMETRY_CONTROL.xSupported OR NOT GVL_GEOMETRY_CONTROL.astStatus[2].xError OR GVL_GEOMETRY_CONTROL.astStatus[2].xResetAllowed)
	AND (NOT GVL_CELL_MANAGER.Status.xError OR GVL_CELL_MANAGER.Status.xResetAllowed)
	AND (NOT GVL_ROBOT.Status.xError OR GVL_ROBOT.Status.xResetAllowed)
	AND (NOT GVL_MACHINE.Status[1].xError OR GVL_MACHINE.Status[1].xResetAllowed)
	AND (NOT GVL_MACHINE.Status[2].xError OR GVL_MACHINE.Status[2].xResetAllowed)
	AND (NOT GVL_MACHINE.Status[3].xError OR GVL_MACHINE.Status[3].xResetAllowed)
	AND (NOT GVL_MAGAZINE.astPartStatus[1].xError
		OR (GVL_MAGAZINE.astError[1].dwAlarmActive = DWORD#0)
		OR fbMagazine1.FaultStatus.xResetAllowed)
	AND (NOT GVL_MAGAZINE.astPartStatus[2].xError
		OR (GVL_MAGAZINE.astError[2].dwAlarmActive = DWORD#0)
		OR fbMagazine2.FaultStatus.xResetAllowed)
	AND (GVL_HMI.xModbusMode OR NOT GVL_AXIS.arrAxis[1].Status.xError OR AXIS_X.FaultStatus.xResetAllowed)
	AND (GVL_HMI.xModbusMode OR NOT GVL_AXIS.arrAxis[2].Status.xError OR AXIS_Y.FaultStatus.xResetAllowed)
	AND (GVL_HMI.xModbusMode OR NOT GVL_AXIS.arrAxis[3].Status.xError OR AXIS_Z.FaultStatus.xResetAllowed)
	AND (GVL_HMI.xModbusMode OR NOT (GVL_AXIS_GROUP.AxisGroup.Status.xLocalError
		OR GVL_AXIS_GROUP.AxisGroup.Status.xLogicalError
		OR GVL_AXIS_GROUP.AxisGroup.Status.xGroupError)
		OR GROUP_XYZ.FaultStatus.xResetAllowed)
	AND (GVL_HMI.xModbusMode OR (GVL_MOTION_MANAGER.stMotionManager.Error.dwAlarmActive = DWORD#0)
		OR GVL_ROBOT.Status.xResetAllowed)
	AND (GVL_HMI.xModbusMode OR (GVL_POINT_MANAGER.PointManager.Error.dwAlarmActive = DWORD#0)
		OR (GVL_ROBOT.Status.xResetAllowed AND ROBOT.FaultStatus.stPoint.xResetAllowed))
	AND (GVL_HMI.xModbusMode OR (GVL_ROBOT.GripperError.dwAlarmActive = DWORD#0)
		OR (GVL_ROBOT.Status.xResetAllowed AND ROBOT.FaultStatus.stGripper.xResetAllowed));

// Два владельца предупреждений используют один источник журнала и общий счётчик.
FOR uiTwin := 1 TO 2 DO
	IF GVL_MAGAZINE.astDiag[uiTwin].stWarning.udiSequence <> audiPartWarningSeen[uiTwin] THEN
		audiPartWarningSeen[uiTwin] := GVL_MAGAZINE.astDiag[uiTwin].stWarning.udiSequence;
		astMagazineWarningMerged[uiTwin].uiCode := GVL_MAGAZINE.astDiag[uiTwin].stWarning.uiCode;
		astMagazineWarningMerged[uiTwin].udiSequence := astMagazineWarningMerged[uiTwin].udiSequence + 1;
	END_IF;
	IF GVL_TWO_PALLET.astDiag[uiTwin].stWarning.udiSequence <> audiTwinWarningSeen[uiTwin] THEN
		audiTwinWarningSeen[uiTwin] := GVL_TWO_PALLET.astDiag[uiTwin].stWarning.udiSequence;
		astMagazineWarningMerged[uiTwin].uiCode := GVL_TWO_PALLET.astDiag[uiTwin].stWarning.uiCode;
		astMagazineWarningMerged[uiTwin].udiSequence := astMagazineWarningMerged[uiTwin].udiSequence + 1;
	END_IF;
END_FOR;

// В журнал передаются все активные ошибки и предупреждения каждого функционального блока.
astAlarmSource[18].eSource := E_ALARM_SOURCE.GEOMETRY_1;
astAlarmSource[19].eSource := E_ALARM_SOURCE.GEOMETRY_2;
FOR uiGeometry := UINT#1 TO UINT#2 DO
	IF GVL_GEOMETRY_CONTROL.xSupported THEN
		astAlarmSource[17 + uiGeometry].dwAlarmActive := GVL_GEOMETRY_CONTROL.astActiveMemory[uiGeometry].dwAlarm;
	ELSE astAlarmSource[17 + uiGeometry].dwAlarmActive := DWORD#0; END_IF;
	astAlarmSource[17 + uiGeometry].xRobotStopRequired := GVL_GEOMETRY_CONTROL.astStatus[uiGeometry].xRobotStopRequired;
	astAlarmSource[17 + uiGeometry].xGlobalError := GVL_CELL_CONTROL.xGlobalError;
	astAlarmSource[17 + uiGeometry].stWarning := GVL_GEOMETRY_CONTROL.astWarning[uiGeometry];
END_FOR;
astAlarmSource[1].eSource := E_ALARM_SOURCE.CELL;
astAlarmSource[1].dwAlarmActive := GVL_CELL_MANAGER.Error.dwAlarmActive;
astAlarmSource[1].xRobotStopRequired := FALSE;
astAlarmSource[1].xGlobalError := GVL_CELL_CONTROL.xGlobalError;
astAlarmSource[1].stWarning := GVL_CELL_MANAGER.Diag.stWarning;

// Каждый владелец сохраняет собственные код и счётчик. Подмена Diag ячейки
// чужим событием приводила к откату на старое предупреждение в следующем скане.
// ALARM_MANAGER регистрирует все три канала независимо под источником CELL.
astAdditionalCellWarning[1] := GVL_MULTI_TYPE.ConfigStatus.stWarning;
astAdditionalCellWarning[2] := GVL_GEOMETRY_CONTROL.stCellWarning;

astAlarmSource[2].eSource := E_ALARM_SOURCE.ROBOT;
astAlarmSource[2].dwAlarmActive := GVL_ROBOT.Error.dwAlarmActive;
astAlarmSource[2].xRobotStopRequired := FALSE;
astAlarmSource[2].xGlobalError := GVL_CELL_CONTROL.xGlobalError;
astAlarmSource[2].stWarning := GVL_ROBOT.Diag.stWarning;

astAlarmSource[3].eSource := E_ALARM_SOURCE.MACHINE_1;
astAlarmSource[3].dwAlarmActive := GVL_MACHINE.Error[1].dwAlarmActive;
astAlarmSource[3].xRobotStopRequired := GVL_MACHINE.Status[1].xCriticalError;
astAlarmSource[3].xGlobalError := GVL_CELL_CONTROL.xGlobalError;
astAlarmSource[3].stWarning := GVL_MACHINE.Diag[1].stWarning;

astAlarmSource[4].eSource := E_ALARM_SOURCE.MACHINE_2;
astAlarmSource[4].dwAlarmActive := GVL_MACHINE.Error[2].dwAlarmActive;
astAlarmSource[4].xRobotStopRequired := GVL_MACHINE.Status[2].xCriticalError;
astAlarmSource[4].xGlobalError := GVL_CELL_CONTROL.xGlobalError;
astAlarmSource[4].stWarning := GVL_MACHINE.Diag[2].stWarning;

astAlarmSource[5].eSource := E_ALARM_SOURCE.MACHINE_3;
astAlarmSource[5].dwAlarmActive := GVL_MACHINE.Error[3].dwAlarmActive;
astAlarmSource[5].xRobotStopRequired := GVL_MACHINE.Status[3].xCriticalError;
astAlarmSource[5].xGlobalError := GVL_CELL_CONTROL.xGlobalError;
astAlarmSource[5].stWarning := GVL_MACHINE.Diag[3].stWarning;

astAlarmSource[6].eSource := E_ALARM_SOURCE.MAGAZINE_LOGIC_1;
astAlarmSource[6].dwAlarmActive := GVL_MAGAZINE.astError[1].dwAlarmActive;
astAlarmSource[6].xRobotStopRequired := GVL_MAGAZINE.astStatus[1].xRobotStopRequired;
astAlarmSource[6].xGlobalError := GVL_CELL_CONTROL.xGlobalError;
astAlarmSource[6].stWarning := astMagazineWarningMerged[1];

astAlarmSource[7].eSource := E_ALARM_SOURCE.MAGAZINE_LOGIC_2;
astAlarmSource[7].dwAlarmActive := GVL_MAGAZINE.astError[2].dwAlarmActive;
astAlarmSource[7].xRobotStopRequired := GVL_MAGAZINE.astStatus[2].xRobotStopRequired;
astAlarmSource[7].xGlobalError := GVL_CELL_CONTROL.xGlobalError;
astAlarmSource[7].stWarning := astMagazineWarningMerged[2];

// Числовые коды 7 и 8 зарезервированы, чтобы старые записи SQLite не начали
// отображаться как аварии осей X/Y после удаления приводов магазинов.
astAlarmSource[8].eSource := E_ALARM_SOURCE.RESERVED_LEGACY_MAGAZINE_AXIS_1;
astAlarmSource[8].dwAlarmActive := DWORD#0;
astAlarmSource[8].xRobotStopRequired := FALSE;
astAlarmSource[8].xGlobalError := GVL_CELL_CONTROL.xGlobalError;
astAlarmSource[8].stWarning.uiCode := UINT#0;
astAlarmSource[8].stWarning.udiSequence := UDINT#0;

astAlarmSource[9].eSource := E_ALARM_SOURCE.RESERVED_LEGACY_MAGAZINE_AXIS_2;
astAlarmSource[9].dwAlarmActive := DWORD#0;
astAlarmSource[9].xRobotStopRequired := FALSE;
astAlarmSource[9].xGlobalError := GVL_CELL_CONTROL.xGlobalError;
astAlarmSource[9].stWarning.uiCode := UINT#0;
astAlarmSource[9].stWarning.udiSequence := UDINT#0;

astAlarmSource[10].eSource := E_ALARM_SOURCE.AXIS_X;
IF GVL_HMI.xModbusMode THEN astAlarmSource[10].dwAlarmActive := DWORD#0;
ELSE astAlarmSource[10].dwAlarmActive := GVL_AXIS.arrAxis[1].Error.dwAlarmActive; END_IF;
astAlarmSource[10].xRobotStopRequired := FALSE;
astAlarmSource[10].xGlobalError := GVL_CELL_CONTROL.xGlobalError;
astAlarmSource[10].stWarning := GVL_AXIS.arrAxis[1].Diag.stWarning;

astAlarmSource[11].eSource := E_ALARM_SOURCE.AXIS_Y;
IF GVL_HMI.xModbusMode THEN astAlarmSource[11].dwAlarmActive := DWORD#0;
ELSE astAlarmSource[11].dwAlarmActive := GVL_AXIS.arrAxis[2].Error.dwAlarmActive; END_IF;
astAlarmSource[11].xRobotStopRequired := FALSE;
astAlarmSource[11].xGlobalError := GVL_CELL_CONTROL.xGlobalError;
astAlarmSource[11].stWarning := GVL_AXIS.arrAxis[2].Diag.stWarning;

astAlarmSource[12].eSource := E_ALARM_SOURCE.AXIS_Z;
IF GVL_HMI.xModbusMode THEN astAlarmSource[12].dwAlarmActive := DWORD#0;
ELSE astAlarmSource[12].dwAlarmActive := GVL_AXIS.arrAxis[3].Error.dwAlarmActive; END_IF;
astAlarmSource[12].xRobotStopRequired := FALSE;
astAlarmSource[12].xGlobalError := GVL_CELL_CONTROL.xGlobalError;
astAlarmSource[12].stWarning := GVL_AXIS.arrAxis[3].Diag.stWarning;

astAlarmSource[13].eSource := E_ALARM_SOURCE.AXIS_GROUP;
IF GVL_HMI.xModbusMode THEN astAlarmSource[13].dwAlarmActive := DWORD#0;
ELSE astAlarmSource[13].dwAlarmActive := GVL_AXIS_GROUP.AxisGroup.Error.dwAlarmActive; END_IF;
astAlarmSource[13].xRobotStopRequired := FALSE;
astAlarmSource[13].xGlobalError := GVL_CELL_CONTROL.xGlobalError;
astAlarmSource[13].stWarning := GVL_AXIS_GROUP.AxisGroup.Diag.stWarning;

astAlarmSource[14].eSource := E_ALARM_SOURCE.MOTION_MANAGER;
IF GVL_HMI.xModbusMode THEN astAlarmSource[14].dwAlarmActive := DWORD#0;
ELSE astAlarmSource[14].dwAlarmActive := GVL_MOTION_MANAGER.stMotionManager.Error.dwAlarmActive; END_IF;
astAlarmSource[14].xRobotStopRequired := FALSE;
astAlarmSource[14].xGlobalError := GVL_CELL_CONTROL.xGlobalError;
astAlarmSource[14].stWarning := GVL_MOTION_MANAGER.stMotionManager.Diag.stWarning;

astAlarmSource[15].eSource := E_ALARM_SOURCE.POINT_MANAGER;
IF GVL_HMI.xModbusMode THEN astAlarmSource[15].dwAlarmActive := DWORD#0;
ELSE astAlarmSource[15].dwAlarmActive := GVL_POINT_MANAGER.PointManager.Error.dwAlarmActive; END_IF;
astAlarmSource[15].xRobotStopRequired := FALSE;
astAlarmSource[15].xGlobalError := GVL_CELL_CONTROL.xGlobalError;
astAlarmSource[15].stWarning := GVL_POINT_MANAGER.PointManager.Diag.stWarning;

astAlarmSource[16].eSource := E_ALARM_SOURCE.GRIPPER;
IF GVL_HMI.xModbusMode THEN astAlarmSource[16].dwAlarmActive := DWORD#0;
ELSE astAlarmSource[16].dwAlarmActive := GVL_ROBOT.GripperError.dwAlarmActive; END_IF;
astAlarmSource[16].xRobotStopRequired := FALSE;
astAlarmSource[16].xGlobalError := GVL_CELL_CONTROL.xGlobalError;
astAlarmSource[16].stWarning := GVL_ROBOT.GripperDiag.stWarning;

astAlarmSource[17].eSource := E_ALARM_SOURCE.CELL_SAFETY;
astAlarmSource[17].dwAlarmActive := CELL_SAFETY.Error.dwAlarmActive;
astAlarmSource[17].xRobotStopRequired := TRUE;
astAlarmSource[17].xGlobalError := CELL_SAFETY.Status.xGlobalError;
astAlarmSource[17].stWarning := CELL_SAFETY.Diag.stWarning;

ALARM_MANAGER(
	xResetWarnings := GVL_ALARM.Command.xResetWarnings,
	astAdditionalCellWarning := astAdditionalCellWarning,
	Sources := astAlarmSource,
	Status => GVL_ALARM.Status,
	Events => GVL_ALARM.Events
);
END_METHOD

METHOD PRIVATE ReadPhysicalInputs
// Единственная страница назначения входов. Сначала фильтры, затем технологические FB.
// Тестовые среды используют модели; сырые входы приводов ГК читает RunGeometryControl.
xPhysicalNormal := GVL_CELL_SETTINGS.eTestEnvironment = E_CELL_TEST_ENVIRONMENT.NORMAL;
GVL_PHYSICAL_IO.xNormalActive := xPhysicalNormal AND GVL_PHYSICAL_IO.xMappingVerified;
xPhysicalInputEnable := GVL_PHYSICAL_IO.xNormalActive;

axPhysicalRaw[1] := GVL_PHYSICAL_IO.xDiMachine1Ready;
axPhysicalRaw[2] := GVL_PHYSICAL_IO.xDiMachine1Alarm;
axPhysicalRaw[3] := GVL_PHYSICAL_IO.xDiMachine1DoorOpen;
axPhysicalRaw[4] := GVL_PHYSICAL_IO.xDiMachine1DoorClosed;
axPhysicalRaw[5] := GVL_PHYSICAL_IO.xDiMachine1HatchLocked;
axPhysicalRaw[6] := GVL_PHYSICAL_IO.xDiMachine1SafetyDoorOpen;
axPhysicalRaw[7] := GVL_PHYSICAL_IO.xDiMachine1SafetyDoorClosed;
axPhysicalRaw[8] := GVL_PHYSICAL_IO.xDiMachine1ChuckClamped;
axPhysicalRaw[9] := GVL_PHYSICAL_IO.xDiMachine1ChuckUnclamped;
axPhysicalRaw[10] := GVL_PHYSICAL_IO.xDiMachine1CycleActive;
axPhysicalRaw[11] := GVL_PHYSICAL_IO.xDiMachine1CycleDone;
axPhysicalRaw[12] := GVL_PHYSICAL_IO.xDiMachine2Ready;
axPhysicalRaw[13] := GVL_PHYSICAL_IO.xDiMachine2Alarm;
axPhysicalRaw[14] := GVL_PHYSICAL_IO.xDiMachine2DoorOpen;
axPhysicalRaw[15] := GVL_PHYSICAL_IO.xDiMachine2DoorClosed;
axPhysicalRaw[16] := GVL_PHYSICAL_IO.xDiMachine2HatchLocked;
axPhysicalRaw[17] := GVL_PHYSICAL_IO.xDiMachine2SafetyDoorOpen;
axPhysicalRaw[18] := GVL_PHYSICAL_IO.xDiMachine2SafetyDoorClosed;
axPhysicalRaw[19] := GVL_PHYSICAL_IO.xDiMachine2ChuckClamped;
axPhysicalRaw[20] := GVL_PHYSICAL_IO.xDiMachine2ChuckUnclamped;
axPhysicalRaw[21] := GVL_PHYSICAL_IO.xDiMachine2CycleActive;
axPhysicalRaw[22] := GVL_PHYSICAL_IO.xDiMachine2CycleDone;
axPhysicalRaw[23] := GVL_PHYSICAL_IO.xDiMachine3Ready;
axPhysicalRaw[24] := GVL_PHYSICAL_IO.xDiMachine3Alarm;
axPhysicalRaw[25] := GVL_PHYSICAL_IO.xDiMachine3DoorOpen;
axPhysicalRaw[26] := GVL_PHYSICAL_IO.xDiMachine3DoorClosed;
axPhysicalRaw[27] := GVL_PHYSICAL_IO.xDiMachine3HatchLocked;
axPhysicalRaw[28] := GVL_PHYSICAL_IO.xDiMachine3SafetyDoorOpen;
axPhysicalRaw[29] := GVL_PHYSICAL_IO.xDiMachine3SafetyDoorClosed;
axPhysicalRaw[30] := GVL_PHYSICAL_IO.xDiMachine3ChuckClamped;
axPhysicalRaw[31] := GVL_PHYSICAL_IO.xDiMachine3ChuckUnclamped;
axPhysicalRaw[32] := GVL_PHYSICAL_IO.xDiMachine3CycleActive;
axPhysicalRaw[33] := GVL_PHYSICAL_IO.xDiMachine3CycleDone;
axPhysicalRaw[34] := GVL_PHYSICAL_IO.xDiGripper1Open;
axPhysicalRaw[35] := GVL_PHYSICAL_IO.xDiGripper1Closed;
axPhysicalRaw[36] := GVL_PHYSICAL_IO.xDiGripper2Open;
axPhysicalRaw[37] := GVL_PHYSICAL_IO.xDiGripper2Closed;
axPhysicalRaw[38] := GVL_PHYSICAL_IO.xDiRotatedToBlank;
axPhysicalRaw[39] := GVL_PHYSICAL_IO.xDiRotatedToDetail;
axPhysicalRaw[40] := GVL_PHYSICAL_IO.xDiCellStartButtonInput;
axPhysicalRaw[41] := GVL_PHYSICAL_IO.xDiCellStopButtonInput;
axPhysicalRaw[42] := GVL_PHYSICAL_IO.xDiCellResetButtonInput;
axPhysicalRaw[43] := GVL_PHYSICAL_IO.xDiEmergencyStopStation1Ok;
axPhysicalRaw[44] := GVL_PHYSICAL_IO.xDiEmergencyStopStation2Ok;
axPhysicalRaw[45] := GVL_PHYSICAL_IO.xDiEmergencyStopStation3Ok;
axPhysicalRaw[46] := GVL_PHYSICAL_IO.xDiEmergencyStopStation4Ok;
axPhysicalRaw[47] := GVL_PHYSICAL_IO.xDiEmergencyStopCabinet1Ok;
axPhysicalRaw[48] := GVL_PHYSICAL_IO.xDiEmergencyStopCabinet2Ok;
axPhysicalRaw[49] := GVL_PHYSICAL_IO.xDiEmergencyStopMpgOk;
axPhysicalRaw[50] := GVL_PHYSICAL_IO.xDiDoor1LockClosed;
axPhysicalRaw[51] := GVL_PHYSICAL_IO.xDiDoor2LockClosed;
axPhysicalRaw[52] := GVL_PHYSICAL_IO.xDiDoor3LockClosed;
axPhysicalRaw[53] := GVL_PHYSICAL_IO.xDiDoor4LockClosed;
axPhysicalRaw[54] := GVL_PHYSICAL_IO.xDiSafetyRelayOkInput;
axPhysicalRaw[55] := GVL_PHYSICAL_IO.xDiPhaseRelayOkInput;
axPhysicalRaw[56] := GVL_PHYSICAL_IO.xDiPressureRelayOkInput;
axPhysicalRaw[57] := GVL_PHYSICAL_IO.xDiMpgAxisXInput;
axPhysicalRaw[58] := GVL_PHYSICAL_IO.xDiMpgAxisYInput;
axPhysicalRaw[59] := GVL_PHYSICAL_IO.xDiMpgAxisZInput;
axPhysicalRaw[60] := GVL_PHYSICAL_IO.xDiMpgMultiplier1Input;
axPhysicalRaw[61] := GVL_PHYSICAL_IO.xDiMpgMultiplier10Input;
axPhysicalRaw[62] := GVL_PHYSICAL_IO.xDiMpgMultiplier100Input;
axPhysicalRaw[63] := GVL_PHYSICAL_IO.xDiMagazine1LockIn;
axPhysicalRaw[64] := GVL_PHYSICAL_IO.xDiMagazine1LockOut;
axPhysicalRaw[65] := GVL_PHYSICAL_IO.xDiMagazine1StopIn;
axPhysicalRaw[66] := GVL_PHYSICAL_IO.xDiMagazine1StopOut;
axPhysicalRaw[67] := GVL_PHYSICAL_IO.xDiMagazine1LiftUp;
axPhysicalRaw[68] := GVL_PHYSICAL_IO.xDiMagazine1LiftDown;
axPhysicalRaw[69] := GVL_PHYSICAL_IO.xDiDoor1UnlockButton;
axPhysicalRaw[70] := GVL_PHYSICAL_IO.xDiDoor2UnlockButton;
axPhysicalRaw[71] := GVL_PHYSICAL_IO.xDiDoor3UnlockButton;
axPhysicalRaw[72] := GVL_PHYSICAL_IO.xDiDoor4UnlockButton;
axPhysicalRaw[73] := GVL_PHYSICAL_IO.xDiMagazine2LockIn;
axPhysicalRaw[74] := GVL_PHYSICAL_IO.xDiMagazine2LockOut;
axPhysicalRaw[75] := GVL_PHYSICAL_IO.xDiMagazine2StopIn;
axPhysicalRaw[76] := GVL_PHYSICAL_IO.xDiMagazine2StopOut;
axPhysicalRaw[77] := GVL_PHYSICAL_IO.xDiMagazine2LiftUp;
axPhysicalRaw[78] := GVL_PHYSICAL_IO.xDiMagazine2LiftDown;

axPhysicalRaw[79] := GVL_PHYSICAL_IO.xDiGk1PartAtEnd;
axPhysicalRaw[80] := GVL_PHYSICAL_IO.xDiGk2PartAtEnd;

axPhysicalRaw[81] := GVL_PHYSICAL_IO.xDiGk1DriveAlarm;
axPhysicalRaw[82] := GVL_PHYSICAL_IO.xDiGk1DriveRunning;
axPhysicalRaw[83] := GVL_PHYSICAL_IO.xDiGk2DriveAlarm;
axPhysicalRaw[84] := GVL_PHYSICAL_IO.xDiGk2DriveRunning;
// Клеммы сохраняются отдельно: ручная подмена не пишет в переменную I/O Mapping.
FOR uiIoIndex := UINT#1 TO UINT#84 DO
    axIoRawDi[uiIoIndex] := axPhysicalRaw[uiIoIndex];
END_FOR;
ReadIoOverrides();
FOR uiIoIndex := UINT#1 TO UINT#84 DO
    IF axIoForced[uiIoIndex] THEN
        axPhysicalRaw[uiIoIndex] := axIoForceValue[uiIoIndex];
    END_IF;
END_FOR;

FOR uiPhysicalInput := 1 TO 80 DO
	tPhysicalRise := GVL_CELL_SETTINGS.tInputFilterRise;
	tPhysicalFall := GVL_CELL_SETTINGS.tInputFilterFall;
	// Срабатывание опасного состояния не задерживается; восстановление фильтруется.
	CASE uiPhysicalInput OF
		2, 13, 24, 41:
			tPhysicalRise := T#0MS;
		1, 3, 4, 5, 6, 7, 8, 9, 12, 14, 15, 16, 17, 18, 19, 20, 23, 25, 26, 27, 28, 29, 30, 31, 34, 35, 36, 37, 38, 39, 43, 44, 45, 46, 47, 48, 49, 50, 51, 52, 53, 54, 55, 56, 63, 64, 65, 66, 67, 68, 73, 74, 75, 76, 77, 78, 79, 80:
			tPhysicalFall := T#0MS;
	END_CASE;
	xPhysicalInputEnable := xPhysicalNormal AND (GVL_PHYSICAL_IO.xMappingVerified OR axIoForced[uiPhysicalInput]);
	afbPhysicalInputFilter[uiPhysicalInput](
		xEnable := xPhysicalInputEnable, xInput := axPhysicalRaw[uiPhysicalInput],
		tRise := tPhysicalRise, tFall := tPhysicalFall);
	axPhysicalFiltered[uiPhysicalInput] := afbPhysicalInputFilter[uiPhysicalInput].xFiltered;
	IF NOT xPhysicalInputEnable THEN
		axPhysicalButtonArmed[uiPhysicalInput] := FALSE;
	ELSIF NOT axPhysicalRaw[uiPhysicalInput] THEN
		axPhysicalButtonArmed[uiPhysicalInput] := TRUE;
	END_IF;
END_FOR;

// Датчики используются FB_GEOMETRY_CONTROL; в NORMAL доступна диагностическая подмена до подтверждения карты.
GVL_PHYSICAL_IO.axGkPartAtEnd[1] := axPhysicalFiltered[79];
GVL_PHYSICAL_IO.axGkPartAtEnd[2] := axPhysicalFiltered[80];

IF xPhysicalNormal THEN
	GVL_MACHINE.astPhysicalInput[1].xReady := axPhysicalFiltered[1];
	GVL_MACHINE.astPhysicalInput[1].xAlarm := axPhysicalFiltered[2];
	GVL_MACHINE.astPhysicalInput[1].xDoorOpen := axPhysicalFiltered[3];
	GVL_MACHINE.astPhysicalInput[1].xDoorClosed := axPhysicalFiltered[4];
	GVL_MACHINE.astPhysicalInput[1].xHatchLocked := axPhysicalFiltered[5];
	GVL_MACHINE.astPhysicalInput[1].xSafetyDoorOpen := axPhysicalFiltered[6];
	GVL_MACHINE.astPhysicalInput[1].xSafetyDoorClosed := axPhysicalFiltered[7];
	GVL_MACHINE.astPhysicalInput[1].xChuckClamped := axPhysicalFiltered[8];
	GVL_MACHINE.astPhysicalInput[1].xChuckUnclamped := axPhysicalFiltered[9];
	GVL_MACHINE.astPhysicalInput[1].xCycleActive := axPhysicalFiltered[10];
	GVL_MACHINE.astPhysicalInput[1].xCycleDone := axPhysicalFiltered[11];
	GVL_MACHINE.astPhysicalInput[2].xReady := axPhysicalFiltered[12];
	GVL_MACHINE.astPhysicalInput[2].xAlarm := axPhysicalFiltered[13];
	GVL_MACHINE.astPhysicalInput[2].xDoorOpen := axPhysicalFiltered[14];
	GVL_MACHINE.astPhysicalInput[2].xDoorClosed := axPhysicalFiltered[15];
	GVL_MACHINE.astPhysicalInput[2].xHatchLocked := axPhysicalFiltered[16];
	GVL_MACHINE.astPhysicalInput[2].xSafetyDoorOpen := axPhysicalFiltered[17];
	GVL_MACHINE.astPhysicalInput[2].xSafetyDoorClosed := axPhysicalFiltered[18];
	GVL_MACHINE.astPhysicalInput[2].xChuckClamped := axPhysicalFiltered[19];
	GVL_MACHINE.astPhysicalInput[2].xChuckUnclamped := axPhysicalFiltered[20];
	GVL_MACHINE.astPhysicalInput[2].xCycleActive := axPhysicalFiltered[21];
	GVL_MACHINE.astPhysicalInput[2].xCycleDone := axPhysicalFiltered[22];
	GVL_MACHINE.astPhysicalInput[3].xReady := axPhysicalFiltered[23];
	GVL_MACHINE.astPhysicalInput[3].xAlarm := axPhysicalFiltered[24];
	GVL_MACHINE.astPhysicalInput[3].xDoorOpen := axPhysicalFiltered[25];
	GVL_MACHINE.astPhysicalInput[3].xDoorClosed := axPhysicalFiltered[26];
	GVL_MACHINE.astPhysicalInput[3].xHatchLocked := axPhysicalFiltered[27];
	GVL_MACHINE.astPhysicalInput[3].xSafetyDoorOpen := axPhysicalFiltered[28];
	GVL_MACHINE.astPhysicalInput[3].xSafetyDoorClosed := axPhysicalFiltered[29];
	GVL_MACHINE.astPhysicalInput[3].xChuckClamped := axPhysicalFiltered[30];
	GVL_MACHINE.astPhysicalInput[3].xChuckUnclamped := axPhysicalFiltered[31];
	GVL_MACHINE.astPhysicalInput[3].xCycleActive := axPhysicalFiltered[32];
	GVL_MACHINE.astPhysicalInput[3].xCycleDone := axPhysicalFiltered[33];
	GVL_PHYSICAL_IO.stGripperFeedback.xGripper1Open := axPhysicalFiltered[34];
	GVL_PHYSICAL_IO.stGripperFeedback.xGripper1Closed := axPhysicalFiltered[35];
	GVL_PHYSICAL_IO.stGripperFeedback.xGripper2Open := axPhysicalFiltered[36];
	GVL_PHYSICAL_IO.stGripperFeedback.xGripper2Closed := axPhysicalFiltered[37];
	GVL_PHYSICAL_IO.stGripperFeedback.xRotatedToBlank := axPhysicalFiltered[38];
	GVL_PHYSICAL_IO.stGripperFeedback.xRotatedToDetail := axPhysicalFiltered[39];
	GVL_CELL_SAFETY_IO.xCellStartButtonInput := axPhysicalFiltered[40] AND axPhysicalButtonArmed[40];
	GVL_CELL_SAFETY_IO.xCellStopButtonInput := axPhysicalFiltered[41];
	GVL_CELL_SAFETY_IO.xCellResetButtonInput := axPhysicalFiltered[42] AND axPhysicalButtonArmed[42];
	GVL_CELL_SAFETY_IO.axEmergencyStopButtonStationInput[1] := NOT axPhysicalFiltered[43];
	GVL_CELL_SAFETY_IO.axEmergencyStopButtonStationInput[2] := NOT axPhysicalFiltered[44];
	GVL_CELL_SAFETY_IO.axEmergencyStopButtonStationInput[3] := NOT axPhysicalFiltered[45];
	GVL_CELL_SAFETY_IO.axEmergencyStopButtonStationInput[4] := NOT axPhysicalFiltered[46];
	GVL_CELL_SAFETY_IO.axEmergencyStopCabinetInput[1] := NOT axPhysicalFiltered[47];
	GVL_CELL_SAFETY_IO.axEmergencyStopCabinetInput[2] := NOT axPhysicalFiltered[48];
	GVL_CELL_SAFETY_IO.xEmergencyStopMpgInput := NOT axPhysicalFiltered[49];
	GVL_CELL_SAFETY_IO.axDoorLockClosedInput[1] := axPhysicalFiltered[50];
	GVL_CELL_SAFETY_IO.axDoorLockClosedInput[2] := axPhysicalFiltered[51];
	GVL_CELL_SAFETY_IO.axDoorLockClosedInput[3] := axPhysicalFiltered[52];
	GVL_CELL_SAFETY_IO.axDoorLockClosedInput[4] := axPhysicalFiltered[53];
	GVL_CELL_SAFETY_IO.xSafetyRelayOkInput := axPhysicalFiltered[54];
	GVL_CELL_SAFETY_IO.xPhaseRelayOkInput := axPhysicalFiltered[55];
	GVL_CELL_SAFETY_IO.xPressureRelayOkInput := axPhysicalFiltered[56];
	GVL_CELL_SAFETY_IO.xMpgAxisXInput := axPhysicalFiltered[57];
	GVL_CELL_SAFETY_IO.xMpgAxisYInput := axPhysicalFiltered[58];
	GVL_CELL_SAFETY_IO.xMpgAxisZInput := axPhysicalFiltered[59];
	GVL_CELL_SAFETY_IO.xMpgMultiplier1Input := axPhysicalFiltered[60];
	GVL_CELL_SAFETY_IO.xMpgMultiplier10Input := axPhysicalFiltered[61];
	GVL_CELL_SAFETY_IO.xMpgMultiplier100Input := axPhysicalFiltered[62];
	GVL_TWO_PALLET.astInput[1].xLockIn := axPhysicalFiltered[63];
	GVL_TWO_PALLET.astInput[1].xLockOut := axPhysicalFiltered[64];
	GVL_TWO_PALLET.astInput[1].xStopIn := axPhysicalFiltered[65];
	GVL_TWO_PALLET.astInput[1].xStopOut := axPhysicalFiltered[66];
	GVL_TWO_PALLET.astInput[1].xLiftUp := axPhysicalFiltered[67];
	GVL_TWO_PALLET.astInput[1].xLiftDown := axPhysicalFiltered[68];
	GVL_CELL_SAFETY_IO.axDoorUnlockButtonInput[1] := axPhysicalFiltered[69] AND axPhysicalButtonArmed[69];
	GVL_CELL_SAFETY_IO.axDoorUnlockButtonInput[2] := axPhysicalFiltered[70] AND axPhysicalButtonArmed[70];
	GVL_CELL_SAFETY_IO.axDoorUnlockButtonInput[3] := axPhysicalFiltered[71] AND axPhysicalButtonArmed[71];
	GVL_CELL_SAFETY_IO.axDoorUnlockButtonInput[4] := axPhysicalFiltered[72] AND axPhysicalButtonArmed[72];
	GVL_TWO_PALLET.astInput[2].xLockIn := axPhysicalFiltered[73];
	GVL_TWO_PALLET.astInput[2].xLockOut := axPhysicalFiltered[74];
	GVL_TWO_PALLET.astInput[2].xStopIn := axPhysicalFiltered[75];
	GVL_TWO_PALLET.astInput[2].xStopOut := axPhysicalFiltered[76];
	GVL_TWO_PALLET.astInput[2].xLiftUp := axPhysicalFiltered[77];
	GVL_TWO_PALLET.astInput[2].xLiftDown := axPhysicalFiltered[78];
	GVL_TWO_PALLET.astInput[1].xIoMapped := GVL_PHYSICAL_IO.xNormalActive;
	GVL_TWO_PALLET.astInput[2].xIoMapped := GVL_PHYSICAL_IO.xNormalActive;
	GVL_MACHINE.astPhysicalInput[1].tRemaining := T#0MS;
	GVL_MACHINE.astPhysicalInput[2].tRemaining := T#0MS;
	GVL_MACHINE.astPhysicalInput[3].tRemaining := T#0MS;
ELSIF xPhysicalWasNormal THEN
	GVL_CELL_SAFETY_IO.xCellStartButtonInput := FALSE;
	GVL_CELL_SAFETY_IO.xCellStopButtonInput := FALSE;
	GVL_CELL_SAFETY_IO.xCellResetButtonInput := FALSE;
	GVL_CELL_SAFETY_IO.axEmergencyStopButtonStationInput[1] := FALSE;
	GVL_CELL_SAFETY_IO.axEmergencyStopButtonStationInput[2] := FALSE;
	GVL_CELL_SAFETY_IO.axEmergencyStopButtonStationInput[3] := FALSE;
	GVL_CELL_SAFETY_IO.axEmergencyStopButtonStationInput[4] := FALSE;
	GVL_CELL_SAFETY_IO.axEmergencyStopCabinetInput[1] := FALSE;
	GVL_CELL_SAFETY_IO.axEmergencyStopCabinetInput[2] := FALSE;
	GVL_CELL_SAFETY_IO.xEmergencyStopMpgInput := FALSE;
	GVL_CELL_SAFETY_IO.axDoorLockClosedInput[1] := TRUE;
	GVL_CELL_SAFETY_IO.axDoorLockClosedInput[2] := TRUE;
	GVL_CELL_SAFETY_IO.axDoorLockClosedInput[3] := TRUE;
	GVL_CELL_SAFETY_IO.axDoorLockClosedInput[4] := TRUE;
	GVL_CELL_SAFETY_IO.xSafetyRelayOkInput := TRUE;
	GVL_CELL_SAFETY_IO.xPhaseRelayOkInput := TRUE;
	GVL_CELL_SAFETY_IO.xPressureRelayOkInput := TRUE;
	GVL_CELL_SAFETY_IO.xMpgAxisXInput := FALSE;
	GVL_CELL_SAFETY_IO.xMpgAxisYInput := FALSE;
	GVL_CELL_SAFETY_IO.xMpgAxisZInput := FALSE;
	GVL_CELL_SAFETY_IO.xMpgMultiplier1Input := FALSE;
	GVL_CELL_SAFETY_IO.xMpgMultiplier10Input := FALSE;
	GVL_CELL_SAFETY_IO.xMpgMultiplier100Input := FALSE;
	GVL_CELL_SAFETY_IO.axDoorUnlockButtonInput[1] := FALSE;
	GVL_CELL_SAFETY_IO.axDoorUnlockButtonInput[2] := FALSE;
	GVL_CELL_SAFETY_IO.axDoorUnlockButtonInput[3] := FALSE;
	GVL_CELL_SAFETY_IO.axDoorUnlockButtonInput[4] := FALSE;
END_IF;
xPhysicalWasNormal := xPhysicalNormal;
END_METHOD

METHOD PRIVATE RecordIoDiagnostics
// Seqlock закрывает весь снимок, включая упаковку масок после добавления событий.
GVL_HMI.udiIoJournalRevision := GVL_HMI.udiIoJournalRevision + UDINT#1;
xIoSnapshotPublishing := TRUE;

axIoOutput[1] := GVL_PHYSICAL_IO.xDoMachine1HatchClosed;
axIoOutput[2] := GVL_PHYSICAL_IO.xDoMachine1HatchUnLock;
axIoOutput[3] := GVL_PHYSICAL_IO.xDoMachine1ClampChuck;
axIoOutput[4] := GVL_PHYSICAL_IO.xDoMachine1UnclampChuck;
axIoOutput[5] := GVL_PHYSICAL_IO.xDoMachine1StartCycle;
axIoOutput[6] := GVL_PHYSICAL_IO.xDoMachine2HatchClosed;
axIoOutput[7] := GVL_PHYSICAL_IO.xDoMachine2HatchUnLock;
axIoOutput[8] := GVL_PHYSICAL_IO.xDoMachine2ClampChuck;
axIoOutput[9] := GVL_PHYSICAL_IO.xDoMachine2UnclampChuck;
axIoOutput[10] := GVL_PHYSICAL_IO.xDoMachine2StartCycle;
axIoOutput[11] := GVL_PHYSICAL_IO.xDoMachine3HatchClosed;
axIoOutput[12] := GVL_PHYSICAL_IO.xDoMachine3HatchUnLock;
axIoOutput[13] := GVL_PHYSICAL_IO.xDoMachine3ClampChuck;
axIoOutput[14] := GVL_PHYSICAL_IO.xDoMachine3UnclampChuck;
axIoOutput[15] := GVL_PHYSICAL_IO.xDoMachine3StartCycle;
axIoOutput[16] := GVL_PHYSICAL_IO.xDoGripper1Open;
axIoOutput[17] := GVL_PHYSICAL_IO.xDoGripper2Open;
axIoOutput[18] := GVL_PHYSICAL_IO.xDoRotateToDetail;
axIoOutput[19] := GVL_PHYSICAL_IO.xDoDoor1Unlock;
axIoOutput[27] := GVL_PHYSICAL_IO.xDoDoor1ButtonLamp;
axIoOutput[20] := GVL_PHYSICAL_IO.xDoDoor2Unlock;
axIoOutput[28] := GVL_PHYSICAL_IO.xDoDoor2ButtonLamp;
axIoOutput[21] := GVL_PHYSICAL_IO.xDoDoor3Unlock;
axIoOutput[29] := GVL_PHYSICAL_IO.xDoDoor3ButtonLamp;
axIoOutput[22] := GVL_PHYSICAL_IO.xDoDoor4Unlock;
axIoOutput[30] := GVL_PHYSICAL_IO.xDoDoor4ButtonLamp;
axIoOutput[23] := GVL_PHYSICAL_IO.xDoSafetyRelayReset;
axIoOutput[24] := GVL_PHYSICAL_IO.xDoSignalTowerGreenOutput;
axIoOutput[25] := GVL_PHYSICAL_IO.xDoSignalTowerAmberOutput;
axIoOutput[26] := GVL_PHYSICAL_IO.xDoSignalTowerRedOutput;
axIoOutput[31] := GVL_PHYSICAL_IO.xDoMagazine1LockIn;
axIoOutput[32] := GVL_PHYSICAL_IO.xDoMagazine1LockOut;
axIoOutput[33] := GVL_PHYSICAL_IO.xDoMagazine1StopIn;
axIoOutput[34] := GVL_PHYSICAL_IO.xDoMagazine1StopOut;
axIoOutput[35] := GVL_PHYSICAL_IO.xDoMagazine1LiftUp;
axIoOutput[36] := GVL_PHYSICAL_IO.xDoMagazine1LiftDown;
axIoOutput[43] := GVL_PHYSICAL_IO.xDoMagazine2LockIn;
axIoOutput[44] := GVL_PHYSICAL_IO.xDoMagazine2LockOut;
axIoOutput[45] := GVL_PHYSICAL_IO.xDoMagazine2StopIn;
axIoOutput[46] := GVL_PHYSICAL_IO.xDoMagazine2StopOut;
axIoOutput[47] := GVL_PHYSICAL_IO.xDoMagazine2LiftUp;
axIoOutput[48] := GVL_PHYSICAL_IO.xDoMagazine2LiftDown;
axIoOutput[37] := FALSE; // Удалённый сигнал; индекс журнала не переиспользовать.
axIoOutput[38] := FALSE; // Удалённый сигнал; индекс журнала не переиспользовать.
axIoOutput[39] := FALSE; // Удалённый сигнал; индекс журнала не переиспользовать.
axIoOutput[40] := GVL_PHYSICAL_IO.xDoCellAlarmHorn;
axIoOutput[41] := GVL_PHYSICAL_IO.xDoGk1DriveRun;
axIoOutput[42] := GVL_PHYSICAL_IO.xDoGk1DriveReset;
axIoOutput[49] := GVL_PHYSICAL_IO.xDoGk2DriveRun;
axIoOutput[50] := GVL_PHYSICAL_IO.xDoGk2DriveReset;
FOR uiIoIndex := UINT#1 TO UINT#80 DO
    axIoUsedDi[uiIoIndex] := axPhysicalFiltered[uiIoIndex];
END_FOR;
FOR uiIoIndex := UINT#81 TO UINT#84 DO
    axIoUsedDi[uiIoIndex] := xPhysicalNormal AND (GVL_PHYSICAL_IO.xMappingVerified OR axIoForced[uiIoIndex]) AND axPhysicalRaw[uiIoIndex];
END_FOR;
FOR uiIoIndex := UINT#1 TO UINT#84 DO
    IF xIoInitialized AND (axIoRawDi[uiIoIndex] <> axIoPreviousRaw[uiIoIndex]) THEN
        AppendIoEvent(usiDirection := USINT#1, uiIndex := uiIoIndex, usiKind := USINT#1,
            xOld := axIoPreviousRaw[uiIoIndex], xNew := axIoRawDi[uiIoIndex]);
    END_IF;
    IF xIoInitialized AND (axIoUsedDi[uiIoIndex] <> axIoPreviousUsed[uiIoIndex]) THEN
        AppendIoEvent(usiDirection := USINT#1, uiIndex := uiIoIndex, usiKind := USINT#2,
            xOld := axIoPreviousUsed[uiIoIndex], xNew := axIoUsedDi[uiIoIndex]);
    END_IF;
    axIoPreviousRaw[uiIoIndex] := axIoRawDi[uiIoIndex];
    axIoPreviousUsed[uiIoIndex] := axIoUsedDi[uiIoIndex];
END_FOR;
FOR uiIoIndex := UINT#1 TO UINT#50 DO
    IF xIoInitialized AND ((uiIoIndex < UINT#37) OR (uiIoIndex > UINT#39)) AND (axIoOutput[uiIoIndex] <> axIoPreviousOutput[uiIoIndex]) THEN
        AppendIoEvent(usiDirection := USINT#2, uiIndex := uiIoIndex, usiKind := USINT#3,
            xOld := axIoPreviousOutput[uiIoIndex], xNew := axIoOutput[uiIoIndex]);
    END_IF;
    axIoPreviousOutput[uiIoIndex] := axIoOutput[uiIoIndex];
END_FOR;
xIoInitialized := TRUE; // Первый снимок — начальный уровень, а не 131 выдуманное переключение.

FOR uiIoWord := UINT#1 TO UINT#3 DO
    GVL_HMI.adwIoRawDi[uiIoWord] := DWORD#0;
    GVL_HMI.adwIoUsedDi[uiIoWord] := DWORD#0;
    GVL_HMI.adwIoForcedDi[uiIoWord] := DWORD#0;
END_FOR;
FOR uiIoWord := UINT#1 TO UINT#2 DO
    GVL_HMI.adwIoDo[uiIoWord] := DWORD#0;
    GVL_HMI.adwIoDoAllowed[uiIoWord] := DWORD#0;
    GVL_HMI.adwIoDoOnAllowed[uiIoWord] := DWORD#0;
    GVL_HMI.adwIoForcedDo[uiIoWord] := DWORD#0;
    GVL_HMI.adwIoInhibitedDo[uiIoWord] := DWORD#0;
END_FOR;
GVL_HMI.uiIoForcedCount := UINT#0;
FOR uiIoIndex := UINT#1 TO UINT#84 DO
    uiIoWord := ((uiIoIndex - UINT#1) / UINT#32) + UINT#1;
    uiIoBit := (uiIoIndex - UINT#1) MOD UINT#32;
    dwIoBit := SHL(DWORD#1, uiIoBit);
    IF axIoRawDi[uiIoIndex] THEN GVL_HMI.adwIoRawDi[uiIoWord] := GVL_HMI.adwIoRawDi[uiIoWord] OR dwIoBit; END_IF;
    IF axIoUsedDi[uiIoIndex] THEN GVL_HMI.adwIoUsedDi[uiIoWord] := GVL_HMI.adwIoUsedDi[uiIoWord] OR dwIoBit; END_IF;
    IF axIoForced[uiIoIndex] THEN
        GVL_HMI.adwIoForcedDi[uiIoWord] := GVL_HMI.adwIoForcedDi[uiIoWord] OR dwIoBit;
        GVL_HMI.uiIoForcedCount := GVL_HMI.uiIoForcedCount + UINT#1;
    END_IF;
END_FOR;
FOR uiIoIndex := UINT#1 TO UINT#50 DO
    uiIoWord := ((uiIoIndex - UINT#1) / UINT#32) + UINT#1;
    uiIoBit := (uiIoIndex - UINT#1) MOD UINT#32;
    dwIoBit := SHL(DWORD#1, uiIoBit);
    IF axIoDoAllowed[uiIoIndex] THEN GVL_HMI.adwIoDoAllowed[uiIoWord] := GVL_HMI.adwIoDoAllowed[uiIoWord] OR dwIoBit; END_IF;
    IF axIoDoOnAllowed[uiIoIndex] THEN GVL_HMI.adwIoDoOnAllowed[uiIoWord] := GVL_HMI.adwIoDoOnAllowed[uiIoWord] OR dwIoBit; END_IF;
    IF axIoDoForced[uiIoIndex] THEN GVL_HMI.adwIoForcedDo[uiIoWord] := GVL_HMI.adwIoForcedDo[uiIoWord] OR dwIoBit; END_IF;
    IF axIoDoInhibited[uiIoIndex] THEN GVL_HMI.adwIoInhibitedDo[uiIoWord] := GVL_HMI.adwIoInhibitedDo[uiIoWord] OR dwIoBit; END_IF;
    IF axIoOutput[uiIoIndex] THEN GVL_HMI.adwIoDo[uiIoWord] := GVL_HMI.adwIoDo[uiIoWord] OR SHL(DWORD#1, uiIoBit); END_IF;
END_FOR;
xIoSnapshotPublishing := FALSE;
GVL_HMI.udiIoJournalRevision := GVL_HMI.udiIoJournalRevision + UDINT#1;
END_METHOD

METHOD PRIVATE PublishGeometryControl
VAR
	uiWarningEvent : UINT;
	xWaitWarningActive : BOOL;
END_VAR
GVL_HMI.astGeometryStatus := GVL_GEOMETRY_CONTROL.astStatus;
// Подсветка следует накопленному предупреждению, включая его сброс в этом скане.
xWaitWarningActive := FALSE;
FOR uiWarningEvent := UINT#1 TO UINT#100 DO
	IF GVL_ALARM.Events[uiWarningEvent].xActive
	AND (GVL_ALARM.Events[uiWarningEvent].eSource = E_ALARM_SOURCE.CELL)
	AND (GVL_ALARM.Events[uiWarningEvent].eSeverity = E_ALARM_SEVERITY.WARNING)
	AND (GVL_ALARM.Events[uiWarningEvent].uiCode = UINT#52) THEN xWaitWarningActive := TRUE; END_IF;
END_FOR;
FOR uiGeometry := UINT#1 TO UINT#2 DO
	GVL_HMI.astGeometryStatus[uiGeometry].xCallWaitWarning := xWaitWarningActive
		AND (GVL_GEOMETRY_CONTROL.astStatus[uiGeometry].xEnabled
			OR NOT (GVL_GEOMETRY_CONTROL.astStatus[1].xEnabled OR GVL_GEOMETRY_CONTROL.astStatus[2].xEnabled));
END_FOR;
GVL_HMI.astGeometryConfig := GVL_GEOMETRY_CONTROL.astActiveConfig;
GVL_HMI.astGeometryCalls := GVL_GEOMETRY_CONTROL.astCalls;
GVL_HMI.auiGeometryPeriod := GVL_GEOMETRY_CONTROL.auiPeriod;
GVL_HMI.auiGeometryCount := GVL_GEOMETRY_CONTROL.auiActiveCount;
GVL_HMI.axGeometryCallAllowed := GVL_GEOMETRY_CONTROL.axCallAllowed;
GVL_HMI.axGeometryCancelAllowed := GVL_GEOMETRY_CONTROL.axCancelAllowed;
GVL_HMI.xGeometryAutoEnabled := GVL_GEOMETRY_CONTROL.xAutoEnabled;
GVL_HMI.xGeometryAutoChangeAllowed := GVL_GEOMETRY_CONTROL.xAutoChangeAllowed;
GVL_HMI.xGeometrySupported := GVL_GEOMETRY_CONTROL.xSupported;
GVL_HMI.xGeometryWaitWhenOccupied := GVL_GEOMETRY_CONTROL.xWaitWhenOccupied;
GVL_HMI.tGeometryTransportTimeout := GVL_GEOMETRY_CONTROL.tTransportTimeout;
GVL_HMI.tGeometryFeedbackTimeout := GVL_GEOMETRY_CONTROL.tDriveFeedbackTimeout;
GVL_HMI.tGeometryResetPulse := GVL_GEOMETRY_CONTROL.tResetPulse;
GVL_HMI.tGeometryWaitWarningTimeout := GVL_GEOMETRY_CONTROL.tWaitWarningTimeout;
GVL_HMI.xGeometrySettingsAllowed := GVL_GEOMETRY_CONTROL.xSettingsAllowed;
// Снимок FIFO имеет версию: gateway читает одинаковый Seq до/после payload.
GVL_HMI.udiGeometryEventSequence := UDINT#0;
GVL_HMI.astGeometryEvents := GVL_GEOMETRY_CONTROL.astEvents;
GVL_HMI.udiGeometryEventSequence := GVL_GEOMETRY_CONTROL.udiEventSequence;
IF GVL_CELL_SETTINGS.eTestEnvironment = E_CELL_TEST_ENVIRONMENT.NORMAL THEN
	GVL_GEOMETRY_CONTROL.astMemory := GVL_GEOMETRY_CONTROL.astActiveMemory;
	GVL_GEOMETRY_CONTROL.astRetainCalls := GVL_GEOMETRY_CONTROL.astCalls;
	GVL_GEOMETRY_CONTROL.auiCount := GVL_GEOMETRY_CONTROL.auiActiveCount;
ELSE
	GVL_GEOMETRY_CONTROL.astSimulationMemory := GVL_GEOMETRY_CONTROL.astActiveMemory;
	GVL_GEOMETRY_CONTROL.astSimulationCalls := GVL_GEOMETRY_CONTROL.astCalls;
	GVL_GEOMETRY_CONTROL.auiSimulationCount := GVL_GEOMETRY_CONTROL.auiActiveCount;
END_IF;
// Фиксированные владельцы счётчиков: переключение среды не меняет идентичность
// OPC UA тега и не превращает старое значение NORMAL в выпуск SIMULATION.
FOR uiGeometry := UINT#1 TO UINT#2 DO
	GVL_HMI.audiGeometryProducedNormal[uiGeometry] := GVL_GEOMETRY_CONTROL.astMemory[uiGeometry].udiProducedPartsTotal;
	GVL_HMI.audiGeometryProducedSimulation[uiGeometry] := GVL_GEOMETRY_CONTROL.astSimulationMemory[uiGeometry].udiProducedPartsTotal;
END_FOR;
END_METHOD

METHOD PRIVATE SetApplicationDefaults
// При старте PLC ячейка всегда включается в ручном режиме: автоматический цикл
// требует явного переключения оператором. Однократный флаг также повторно
// применяет безопасные значения при Online Change, когда initializer GVL
// может не перезаписать уже существующее значение. Инициализация выполняется до
// RunCellControl, чтобы автомат не увидел прежние настройки даже на один цикл.
IF NOT xApplicationStartupInitialized THEN
	GVL_CELL_CONTROL.xManual := TRUE;
	FOR uiMachine := 1 TO 3 DO
		GVL_HMI.axMachineUsed[uiMachine] := FALSE;
	END_FOR;
	// RETAIN uiMode переживает перезапуск PLC, поэтому явно выбираем двухпалетный
	// тип на старте. При реальной смене типа старые базы магазинов недействительны.
	IF GVL_TWO_PALLET.uiMode <> UINT#1 THEN
		GVL_TWO_PALLET.uiMode := UINT#1;
		GVL_POINT.astRetainPoints[UINT#14].xConfigured := FALSE;
		GVL_POINT.astRetainPoints[UINT#15].xConfigured := FALSE;
		xPointTableReady := FALSE;
	END_IF;
	GVL_CELL_SETTINGS.eTestEnvironment := E_CELL_TEST_ENVIRONMENT.SIMULATION;
	xApplicationStartupInitialized := TRUE;
END_IF;

// При первом запуске этой схемы намеренно отбрасываем прежние инженерные
// координаты. Нулевая скорость и xConfigured=FALSE не позволяют принять
// нулевую точку за пригодную для движения.
IF GVL_POINT.udiPointStorageVersion <> GVL_POINT.udiExpectedPointStorageVersion THEN
	FOR uiPointEditorIndex := UINT#1 TO INT_TO_UINT(GVL_POINT.iPersistentPointCapacity) DO
		GVL_POINT.astRetainPoints[uiPointEditorIndex].Name := '';
		GVL_POINT.astRetainPoints[uiPointEditorIndex].X := 0.0;
		GVL_POINT.astRetainPoints[uiPointEditorIndex].Y := 0.0;
		GVL_POINT.astRetainPoints[uiPointEditorIndex].Z := 0.0;
		GVL_POINT.astRetainPoints[uiPointEditorIndex].MagazineSafeZ := 0.0;
		GVL_POINT.astRetainPoints[uiPointEditorIndex].MagazineChangeZ := 0.0;
		GVL_POINT.astRetainPoints[uiPointEditorIndex].SpeedFactor := 0.0;
		GVL_POINT.astRetainPoints[uiPointEditorIndex].xConfigured := FALSE;
	END_FOR;
	GVL_POINT.udiPointStorageVersion := GVL_POINT.udiExpectedPointStorageVersion;
END_IF;

// Единственное соответствие компактного редакторского индекса, стабильного
// E_POINT_NAME и прежнего индекса Persistent-массива. Три legacy-точки INSIDE
// пропущены; рецепты станков их не используют.
xPointTableReady := TRUE;
// Базы ГК хранятся у владельца GVL_GEOMETRY_CONTROL, отдельно от прежних 15
// Persistent-позиций. Их добавление не сбрасывает уже сохранённые точки.
FOR uiPointEditorIndex := UINT#1 TO INT_TO_UINT(GVL_POINT.iRequiredPointCount) DO
	uiPointStorageIndex := UINT#0;
	CASE uiPointEditorIndex OF
		UINT#1: ePointEditorName := E_POINT_NAME.MACHINE_1_ABOVE; uiPointStorageIndex := UINT#1;
		UINT#2: ePointEditorName := E_POINT_NAME.MACHINE_1_CHUCK_APROACH; uiPointStorageIndex := UINT#3;
		UINT#3: ePointEditorName := E_POINT_NAME.MACHINE_1_CHUCK_POSITION; uiPointStorageIndex := UINT#4;
		UINT#4: ePointEditorName := E_POINT_NAME.MACHINE_2_ABOVE; uiPointStorageIndex := UINT#5;
		UINT#5: ePointEditorName := E_POINT_NAME.MACHINE_2_CHUCK_APROACH; uiPointStorageIndex := UINT#7;
		UINT#6: ePointEditorName := E_POINT_NAME.MACHINE_2_CHUCK_POSITION; uiPointStorageIndex := UINT#8;
		UINT#7: ePointEditorName := E_POINT_NAME.MACHINE_3_ABOVE; uiPointStorageIndex := UINT#9;
		UINT#8: ePointEditorName := E_POINT_NAME.MACHINE_3_CHUCK_APROACH; uiPointStorageIndex := UINT#11;
		UINT#9: ePointEditorName := E_POINT_NAME.MACHINE_3_CHUCK_POSITION; uiPointStorageIndex := UINT#12;
		UINT#10: ePointEditorName := E_POINT_NAME.HOME_SAFETY; uiPointStorageIndex := UINT#13;
		UINT#11: ePointEditorName := E_POINT_NAME.MAGAZINE_1_DETAIL; uiPointStorageIndex := UINT#14;
		UINT#12: ePointEditorName := E_POINT_NAME.MAGAZINE_2_DETAIL; uiPointStorageIndex := UINT#15;
	ELSE
		ePointEditorName := E_POINT_NAME.NONE;
	END_CASE;

	IF (ePointEditorName <> E_POINT_NAME.NONE) AND (uiPointStorageIndex <> UINT#0) THEN
		GVL_POINT.Points[ePointEditorName] := GVL_POINT.astRetainPoints[uiPointStorageIndex];
		IF (ePointEditorName = E_POINT_NAME.MAGAZINE_1_DETAIL)
		OR (ePointEditorName = E_POINT_NAME.MAGAZINE_2_DETAIL) THEN
			GVL_POINT.Points[ePointEditorName].xConfigured :=
				GVL_POINT.astRetainPoints[uiPointStorageIndex].xConfigured
				AND (GVL_POINT.astRetainPoints[uiPointStorageIndex].MagazineSafeZ <> LREAL#0.0)
				AND (GVL_POINT.astRetainPoints[uiPointStorageIndex].MagazineChangeZ <> LREAL#0.0);
		END_IF;
		IF NOT GVL_POINT.Points[ePointEditorName].xConfigured THEN
			xPointTableReady := FALSE;
		END_IF;
	ELSE
		xPointTableReady := FALSE;
	END_IF;
END_FOR;

// Полнота таблицы остаётся диагностикой редактора. Включение оборудования
// проверяет только собственные точки; HOME_SAFETY отдельно нужен автоциклу.
axMachinePointsReady[1] := GVL_POINT.Points[E_POINT_NAME.MACHINE_1_ABOVE].xConfigured
	AND GVL_POINT.Points[E_POINT_NAME.MACHINE_1_CHUCK_APROACH].xConfigured
	AND GVL_POINT.Points[E_POINT_NAME.MACHINE_1_CHUCK_POSITION].xConfigured;
axMachinePointsReady[2] := GVL_POINT.Points[E_POINT_NAME.MACHINE_2_ABOVE].xConfigured
	AND GVL_POINT.Points[E_POINT_NAME.MACHINE_2_CHUCK_APROACH].xConfigured
	AND GVL_POINT.Points[E_POINT_NAME.MACHINE_2_CHUCK_POSITION].xConfigured;
axMachinePointsReady[3] := GVL_POINT.Points[E_POINT_NAME.MACHINE_3_ABOVE].xConfigured
	AND GVL_POINT.Points[E_POINT_NAME.MACHINE_3_CHUCK_APROACH].xConfigured
	AND GVL_POINT.Points[E_POINT_NAME.MACHINE_3_CHUCK_POSITION].xConfigured;
axMagazinePointsReady[1] := GVL_POINT.Points[E_POINT_NAME.MAGAZINE_1_DETAIL].xConfigured;
axMagazinePointsReady[2] := GVL_POINT.Points[E_POINT_NAME.MAGAZINE_2_DETAIL].xConfigured;
END_METHOD

METHOD PRIVATE RunSafety
FOR uiTwin := 1 TO 2 DO
	axTwinSafetyBusy[uiTwin] := (GVL_TWO_PALLET.uiMode = 1) AND (GVL_TWO_PALLET.astStatus[uiTwin].xBusy
		OR (GVL_TWO_PALLET.astInput[uiTwin].xAxisBound AND NOT GVL_TWO_PALLET.astInput[uiTwin].xStandstill));
END_FOR;
FOR uiMachine := UINT#1 TO UINT#4 DO
	axButtonStationInput[uiMachine] := GVL_CELL_SAFETY_IO.axDoorUnlockButtonInput[uiMachine]
		OR ((GVL_CELL_SETTINGS.eTestEnvironment = E_CELL_TEST_ENVIRONMENT.SIMULATION)
			AND GVL_CELL_SAFETY_IO.axSimDoorUnlockButtonInput[uiMachine]);
	axButtonStationEmergencyStopInput[uiMachine] := GVL_CELL_SAFETY_IO.axEmergencyStopButtonStationInput[uiMachine]
		OR ((GVL_CELL_SETTINGS.eTestEnvironment = E_CELL_TEST_ENVIRONMENT.SIMULATION)
			AND GVL_CELL_SAFETY_IO.axSimEmergencyStopButtonStationInput[uiMachine]);
END_FOR;
CELL_SAFETY(
	axMagazineMechanismBusy := axTwinSafetyBusy,
	axDoorLockClosedInput := GVL_CELL_SAFETY_IO.axDoorLockClosedInput,
	axDoorUnlockButtonInput := axButtonStationInput,
	axEmergencyStopButtonStationInput := axButtonStationEmergencyStopInput,
	axEmergencyStopCabinetInput := GVL_CELL_SAFETY_IO.axEmergencyStopCabinetInput,
	xEmergencyStopMpgInput := GVL_CELL_SAFETY_IO.xEmergencyStopMpgInput,
	xPhaseRelayOkInput := GVL_CELL_SAFETY_IO.xPhaseRelayOkInput,
	xPressureRelayOkInput := GVL_CELL_SAFETY_IO.xPressureRelayOkInput,
	xSafetyRelayOkInput := GVL_CELL_SAFETY_IO.xSafetyRelayOkInput,
	xCellStartButtonInput := GVL_CELL_SAFETY_IO.xCellStartButtonInput,
	xCellStopButtonInput := GVL_CELL_SAFETY_IO.xCellStopButtonInput,
	xCellResetButtonInput := GVL_CELL_SAFETY_IO.xCellResetButtonInput,
	xMpgAxisXInput := GVL_CELL_SAFETY_IO.xMpgAxisXInput,
	xMpgAxisYInput := GVL_CELL_SAFETY_IO.xMpgAxisYInput,
	xMpgAxisZInput := GVL_CELL_SAFETY_IO.xMpgAxisZInput,
	xMpgMultiplier1Input := GVL_CELL_SAFETY_IO.xMpgMultiplier1Input,
	xMpgMultiplier10Input := GVL_CELL_SAFETY_IO.xMpgMultiplier10Input,
	xMpgMultiplier100Input := GVL_CELL_SAFETY_IO.xMpgMultiplier100Input,
	xSafetyRelayReset := GVL_HMI.xSafetyRelayReset,
	astMagazineStatus := GVL_MAGAZINE.astStatus,
	FaultRequest := stSafetyFaultRequest
);

GVL_CELL_SAFETY_IO.axDoorUnlockOutput := CELL_SAFETY.axDoorUnlockOutput;
GVL_CELL_SAFETY_IO.axDoorButtonLampOutput := CELL_SAFETY.axDoorButtonLampOutput;
GVL_CELL_SAFETY_IO.xSafetyRelayResetOutput := CELL_SAFETY.xSafetyRelayResetOutput;

// Физические Старт/Стоп/Сброс — равноправные дубли HMI-команд, но только по фронту.
GVL_CELL_CONTROL.xEnable := GVL_CELL_CONTROL.xEnable OR CELL_SAFETY.xCellEnablePulse;
GVL_CELL_CONTROL.xDisable := GVL_CELL_CONTROL.xDisable OR CELL_SAFETY.xCellDisablePulse;
GVL_CELL_CONTROL.xReset := GVL_CELL_CONTROL.xReset OR CELL_SAFETY.xCellResetPulse;

// Ручное I/O владеет механизмами. Физический Start также не возобновляет
// прерванный автомат; выход из этого режима сам по себе ничего не запускает.
IF xIoManualActive THEN
	GVL_CELL_CONTROL.xStart := FALSE;
	GVL_CELL_CONTROL.xEnable := FALSE;
	GVL_CELL_CONTROL.xStop := TRUE;
END_IF;

GVL_CELL_CONTROL.xGlobalError := CELL_SAFETY.Status.xGlobalError;

// HMI записывает payload, затем CommandSeq. Gateway удерживает единственного
// писателя до AckSeq. Даже запись между RunSafety и PublishHmi не теряется:
// PLC никогда не перезаписывает запрос, а обработает его в следующем скане.
uiCellModeRejectReason := UINT#0;
udiCellModeCommandSnapshot := GVL_HMI.udiCellModeCommandSeq;
IF (udiCellModeCommandSnapshot <> UDINT#0)
AND (udiCellModeCommandSnapshot <> GVL_HMI.udiCellModeAckSeq) THEN
	IF GVL_HMI.xCellManualRequest
	AND GVL_CELL_MANAGER.Status.xRunning
	AND NOT GVL_CELL_CONTROL.xGlobalError THEN
		uiCellModeRejectReason := UINT#2;
	ELSIF NOT GVL_HMI.xCellManualRequest
	AND (GVL_CELL_CONTROL.xGlobalError OR GVL_HMI.xIoEmergencyStopActive) THEN
		uiCellModeRejectReason := UINT#3;
	ELSE
		GVL_CELL_CONTROL.xManual := GVL_HMI.xCellManualRequest;
	END_IF;
	IF uiCellModeRejectReason = UINT#0 THEN
		GVL_HMI.uiCellModeResult := UINT#1;
	ELSE
		GVL_HMI.uiCellModeResult := uiCellModeRejectReason;
	END_IF;
	// Ack публикуется после фактического режима в PublishHmi, включая отказ.
END_IF;

IF GVL_CELL_CONTROL.xGlobalError OR GVL_HMI.xIoEmergencyStopActive THEN
	GVL_CELL_CONTROL.xManual := TRUE;
END_IF;

// Разрешения рассчитываются после применения режима и Safety текущего скана.
xRobotHmiPermit := GVL_CELL_CONTROL.xManual AND NOT GVL_CELL_MANAGER.Status.xRunning
    AND NOT xIoManualActive
    AND NOT GVL_HMI.xIoEmergencyStopActive;
xRobotAutoPowerOff := NOT GVL_CELL_CONTROL.xManual
	AND (GVL_ROBOT.Status.xError
		OR GVL_AXIS.arrAxis[1].Status.xError
		OR GVL_AXIS.arrAxis[2].Status.xError
		OR GVL_AXIS.arrAxis[3].Status.xError
		OR GVL_AXIS_GROUP.AxisGroup.Status.xLocalError
		OR GVL_AXIS_GROUP.AxisGroup.Status.xLogicalError
		OR GVL_AXIS_GROUP.AxisGroup.Status.xGroupError);
END_METHOD

METHOD PRIVATE ReadIoOverrides
udiIoNowMs := TIME_TO_UDINT(TIME());
IF NOT xIoInitialized THEN
    GVL_HMI.udiIoBootCounter := GVL_HMI.udiIoBootCounter + UDINT#1;
    IF GVL_HMI.udiIoBootCounter = UDINT#0 THEN GVL_HMI.udiIoBootCounter := UDINT#1; END_IF;
    udiIoLastTickMs := udiIoNowMs;
    // Старый запрос после перезапуска не должен исполняться сам собой.
    GVL_HMI.udiIoOverrideAckSeq := GVL_HMI.udiIoOverrideCommandSeq;
    GVL_HMI.udiIoEmergencyAckSeq := GVL_HMI.udiIoEmergencyCommandSeq;
END_IF;
IF udiIoNowMs >= udiIoLastTickMs THEN
    uliIoClockMs := uliIoClockMs + UDINT_TO_ULINT(udiIoNowMs - udiIoLastTickMs);
ELSE
    uliIoClockMs := uliIoClockMs + ULINT#4294967296 - UDINT_TO_ULINT(udiIoLastTickMs) + UDINT_TO_ULINT(udiIoNowMs);
END_IF;
udiIoLastTickMs := udiIoNowMs;
GVL_HMI.sIoClockMs := ULINT_TO_STRING(uliIoClockMs);

tonIoOverrideWatchdog(IN := GVL_HMI.udiIoOverrideHeartbeat = udiIoHeartbeatSeen, PT := T#3S);
IF GVL_HMI.udiIoOverrideHeartbeat <> udiIoHeartbeatSeen THEN
    udiIoHeartbeatSeen := GVL_HMI.udiIoOverrideHeartbeat;
END_IF;
IF udiIoNowMs >= GVL_HMI.udiIoOverrideHeartbeatAtMs THEN
    uliIoLeaseAgeMs := UDINT_TO_ULINT(udiIoNowMs) - UDINT_TO_ULINT(GVL_HMI.udiIoOverrideHeartbeatAtMs);
ELSE
    uliIoLeaseAgeMs := ULINT#4294967296 + UDINT_TO_ULINT(udiIoNowMs) - UDINT_TO_ULINT(GVL_HMI.udiIoOverrideHeartbeatAtMs);
END_IF;

xIoBusy := GVL_CELL_MANAGER.Status.xRunning OR GVL_CELL_MANAGER.Status.xBusy
    OR GVL_CELL_MANAGER.Status.xStopPending OR GVL_ROBOT.Status.xBusy
    OR xMotionBusy OR xGroupMotionBusy OR xPointCheckActive OR xPointCheckRequest
    OR xPowerTransitionActive OR SIMULATION_DYNAMICS.xBusy
    OR GVL_HMI.xRobotManualExecute OR GVL_HMI.stRobotCommand.xExecute
    OR GVL_CELL_CONTROL.xStart
    OR (GVL_HMI.udiTwinCommandSeq <> GVL_HMI.udiTwinAckSeq);
// Реальный цикл станка нельзя скрыть подменой его DI.
IF xPhysicalNormal AND GVL_PHYSICAL_IO.xMappingVerified THEN
    xIoBusy := xIoBusy OR GVL_PHYSICAL_IO.xDiMachine1CycleActive
        OR GVL_PHYSICAL_IO.xDiMachine2CycleActive OR GVL_PHYSICAL_IO.xDiMachine3CycleActive;
END_IF;
FOR uiIoIndex := UINT#1 TO UINT#3 DO
    xIoBusy := xIoBusy OR GVL_MACHINE.Status[uiIoIndex].xBusy OR GVL_MACHINE.Status[uiIoIndex].xProcessing
        OR GVL_HMI.axMachineManualHatchOpen[uiIoIndex] OR GVL_HMI.axMachineManualHatchClose[uiIoIndex]
        OR GVL_HMI.axMachineManualHatchUnlock[uiIoIndex] OR GVL_HMI.axMachineManualHatchLock[uiIoIndex]
        OR GVL_HMI.axMachineManualChuckOpen[uiIoIndex] OR GVL_HMI.axMachineManualChuckClose[uiIoIndex]
        OR GVL_HMI.astAxisHmiCommand[uiIoIndex].xJogPositive
        OR GVL_HMI.astAxisHmiCommand[uiIoIndex].xJogNegative
        OR GVL_HMI.astAxisHmiCommand[uiIoIndex].xHome
        OR GVL_HMI.astAxisHmiCommand[uiIoIndex].xMoveAbsolute
        OR GVL_HMI.astAxisHmiCommand[uiIoIndex].xMoveRelative;
END_FOR;
FOR uiIoIndex := UINT#1 TO UINT#2 DO
    xIoBusy := xIoBusy OR GVL_MAGAZINE.astStatus[uiIoIndex].xBusy
        OR GVL_TWO_PALLET.astStatus[uiIoIndex].xBusy;
END_FOR;
// Ручной режим сигналов включается одним запросом. Технологических допусков здесь нет.
xIoManualEndedByOperator := FALSE;
IF xIoManualActive AND (NOT GVL_CELL_CONTROL.xManual OR NOT xHmiConnectionAlive
    OR tonIoOverrideWatchdog.Q OR (uliIoLeaseAgeMs > ULINT#3000)
    OR ((GVL_HMI.udiCellModeCommandSeq <> GVL_HMI.udiCellModeAckSeq) AND NOT GVL_HMI.xCellManualRequest)) THEN
    xIoManualActive := FALSE;
END_IF;
// Прямой ручной слой доступен и при зависших Busy/Processing владельцев.
// Их задания отменяются при передаче управления; xIoBusy остаётся диагностикой
// и условием снятия отдельного программного аварийного останова.
GVL_HMI.xIoManualStartAllowed := GVL_CELL_CONTROL.xManual AND NOT xIoManualActive
    AND NOT ((GVL_HMI.udiCellModeCommandSeq <> GVL_HMI.udiCellModeAckSeq) AND NOT GVL_HMI.xCellManualRequest);
xIoOverrideRejected := FALSE;
udiIoRequestSeq := GVL_HMI.udiIoOverrideCommandSeq;
uiIoRequestAction := GVL_HMI.uiIoOverrideAction;
uiIoRequestIndex := GVL_HMI.uiIoOverrideIndex;
xIoRequestValue := GVL_HMI.xIoOverrideValue;
IF udiIoRequestSeq <> GVL_HMI.udiIoOverrideAckSeq THEN
    IF (uiIoRequestAction = UINT#8) OR (uiIoRequestAction = UINT#9) OR (uiIoRequestAction = UINT#7) THEN
        GVL_HMI.uiIoOverrideResult := UINT#4;
        IF IsHmiCommandFresh(udiIssuedAtMs := GVL_HMI.udiIoOverrideIssuedAtMs) THEN
            GVL_HMI.uiIoOverrideResult := UINT#1;
            IF uiIoRequestAction = UINT#8 THEN
                IF NOT xHmiConnectionAlive OR tonIoOverrideWatchdog.Q OR (uliIoLeaseAgeMs > ULINT#3000) THEN
                    GVL_HMI.uiIoOverrideResult := UINT#4;
                ELSIF xIoManualActive THEN
                    // Повтор входа не перезаписывает уже выбранные ручные уровни.
                    GVL_HMI.uiIoOverrideResult := UINT#1;
                ELSIF GVL_HMI.xIoManualStartAllowed THEN
                    FOR uiIoIndex := UINT#1 TO UINT#50 DO
                        axIoDoForceValue[uiIoIndex] := axIoOutput[uiIoIndex];
                        axIoDoForced[uiIoIndex] := FALSE;
                    END_FOR;
                    xIoManualActive := TRUE;
                ELSE
                    GVL_HMI.uiIoOverrideResult := UINT#2;
                END_IF;
            ELSE
                xIoManualActive := FALSE;
                xIoManualEndedByOperator := TRUE;
            END_IF;
        END_IF;
        // Для входа/выхода из режима Ack выдаёт ApplyIoOutputOverrides после назначения DO.
    END_IF;
END_IF;

GVL_HMI.xIoManualControlActive := xIoManualActive;
GVL_HMI.xIoManualStartAllowed := GVL_HMI.xIoManualStartAllowed AND NOT xIoManualActive;
GVL_HMI.xIoOverrideAllowed := xIoManualActive AND GVL_CELL_CONTROL.xManual;
IF GVL_HMI.xIoOverrideAllowed THEN GVL_HMI.uiIoOverrideBlockReason := UINT#0;
ELSIF NOT GVL_CELL_CONTROL.xManual THEN GVL_HMI.uiIoOverrideBlockReason := UINT#2;
ELSE GVL_HMI.uiIoOverrideBlockReason := UINT#7;
END_IF;

IF NOT GVL_HMI.xIoOverrideAllowed THEN
    FOR uiIoIndex := UINT#1 TO UINT#84 DO
        IF axIoForced[uiIoIndex] THEN
            IF xIoManualEndedByOperator THEN
                AppendIoEvent(usiDirection := USINT#1, uiIndex := uiIoIndex, usiKind := USINT#5,
                    xOld := axIoForceValue[uiIoIndex], xNew := axIoRawDi[uiIoIndex]);
            ELSE
                AppendIoEvent(usiDirection := USINT#1, uiIndex := uiIoIndex, usiKind := USINT#6,
                    xOld := axIoForceValue[uiIoIndex], xNew := axIoRawDi[uiIoIndex]);
            END_IF;
            axIoForced[uiIoIndex] := FALSE;
        END_IF;
    END_FOR;
END_IF;

IF (udiIoRequestSeq <> GVL_HMI.udiIoOverrideAckSeq)
AND NOT ((uiIoRequestAction >= UINT#4) AND (uiIoRequestAction <= UINT#9)) THEN
    GVL_HMI.uiIoOverrideResult := UINT#3;
    IF NOT IsHmiCommandFresh(udiIssuedAtMs := GVL_HMI.udiIoOverrideIssuedAtMs) THEN
        GVL_HMI.uiIoOverrideResult := UINT#4;
    ELSIF uiIoRequestAction = UINT#3 THEN
        FOR uiIoIndex := UINT#1 TO UINT#84 DO
            IF axIoForced[uiIoIndex] THEN
                AppendIoEvent(usiDirection := USINT#1, uiIndex := uiIoIndex, usiKind := USINT#5,
                    xOld := axIoForceValue[uiIoIndex], xNew := axIoRawDi[uiIoIndex]);
                axIoForced[uiIoIndex] := FALSE;
            END_IF;
        END_FOR;
        GVL_HMI.uiIoOverrideResult := UINT#1;
    ELSIF (uiIoRequestIndex >= UINT#1) AND (uiIoRequestIndex <= UINT#84) THEN
        IF uiIoRequestAction = UINT#2 THEN
            IF axIoForced[uiIoRequestIndex] THEN
                AppendIoEvent(usiDirection := USINT#1, uiIndex := uiIoRequestIndex, usiKind := USINT#5,
                    xOld := axIoForceValue[uiIoRequestIndex], xNew := axIoRawDi[uiIoRequestIndex]);
                axIoForced[uiIoRequestIndex] := FALSE;
            END_IF;
            GVL_HMI.uiIoOverrideResult := UINT#1;
        ELSIF uiIoRequestAction = UINT#1 THEN
            IF GVL_HMI.xIoOverrideAllowed THEN
                IF NOT axIoForced[uiIoRequestIndex] OR (axIoForceValue[uiIoRequestIndex] <> xIoRequestValue) THEN
                    AppendIoEvent(usiDirection := USINT#1, uiIndex := uiIoRequestIndex, usiKind := USINT#4,
                        xOld := axPhysicalRaw[uiIoRequestIndex], xNew := xIoRequestValue);
                END_IF;
                axIoForced[uiIoRequestIndex] := TRUE;
                axIoForceValue[uiIoRequestIndex] := xIoRequestValue;
                GVL_HMI.uiIoOverrideResult := UINT#1;
            ELSE
                GVL_HMI.uiIoOverrideResult := UINT#2;
            END_IF;
        END_IF;
    END_IF;
    xIoOverrideRejected := GVL_HMI.uiIoOverrideResult <> UINT#1;
    GVL_HMI.udiIoOverrideAckSeq := udiIoRequestSeq;
END_IF;
FOR uiIoIndex := UINT#1 TO UINT#84 DO
    IF axIoForced[uiIoIndex] THEN axPhysicalRaw[uiIoIndex] := axIoForceValue[uiIoIndex]; END_IF;
END_FOR;
END_METHOD

